(* IEC 61131-3 sources: daoli-st-library/DL_Motion (part 16) *)

(* ---- FB_DL_ResolverAngleTrackObs.st ---- *)
(* ===========================================================================
   组件名   : FB_DL_ResolverAngleTrackObs
   分类     : DL_Motion / 旋转变压器角度跟踪观测器
   一句话   : 二阶跟踪环由 sin/cos 直接跟踪角度与转速，无需反三角运算且天然解卷绕
   复杂度   : 3        版本 : v1.0.0        日期 : 2026-11-24
   开源溯源 : 无（clean-room 自研，未借鉴任何开源实现）
   输入契约 : fSin/fCos 两路瞬时值 [V]；fKp 角度环增益 [1/s]；fKi 速度环增益 [1/s²]
              fDtSec 采样周期 [s]；fAmpMin 最小有效幅值 [V]；fSpeedMax 转速限幅 [rad/s]
              fLockBand 锁定判定带宽（归一化误差） | lock band
   输出契约 : fAngleEst 跟踪角 [rad] 0..2π；fSpeedEst 跟踪转速 [rad/s]
              fErrorNorm 归一化角度误差（≈sin(θin−θest)） | normalized angle error
              xLocked 已锁定；xValid 输入有效；eStateOut 状态观测
   修改记录 : v1.0.0 2026-11-24 初版
   =========================================================================== *)

TYPE E_DL_TrackState :
(
    eTrackInit := 0,     // 初始化（粗定位） | init by coarse seed
    eTracking := 1,      // 正常跟踪 | normal tracking
    eSignalLost := 2     // 信号丢失冻结 | signal lost freeze
);
END_TYPE

FUNCTION_BLOCK FB_DL_ResolverAngleTrackObs
VAR_INPUT
    fSin : REAL;                        // 正弦路瞬时值 [V] | sine channel value [V]
    fCos : REAL;                        // 余弦路瞬时值 [V] | cosine channel value [V]
    fKp : REAL := 60.0;                 // 角度环增益 [1/s] | angle loop gain [1/s]
    fKi : REAL := 2000.0;               // 速度环增益 [1/s²] | speed loop gain [1/s^2]
    fDtSec : REAL := 0.0001;            // 采样周期 [s] | sample period [s]
    fAmpMin : REAL := 0.5;              // 最小有效幅值 [V] | minimum valid amplitude [V]
    fSpeedMax : REAL := 500.0;          // 转速限幅 [rad/s] | speed clamp [rad/s]
    fLockBand : REAL := 0.02;           // 锁定判定带宽（归一化） | lock band normalized
END_VAR
VAR_OUTPUT
    fAngleEst : REAL;                   // 跟踪角度 [rad] 0..2π | estimated angle [rad]
    fSpeedEst : REAL;                   // 跟踪转速 [rad/s] | estimated speed [rad/s]
    fErrorNorm : REAL;                  // 归一化角度误差 | normalized angle error
    xLocked : BOOL;                     // 已锁定标志 | locked flag
    xValid : BOOL;                      // 输入有效标志 | inputs valid flag
    eStateOut : E_DL_TrackState;        // 当前状态观测 | current state observation
END_VAR
VAR
    _eState : E_DL_TrackState := eTrackInit;  // 内部状态机状态 | internal state
    _fAngle : REAL;                     // 内部跟踪角 [rad] | internal tracked angle [rad]
    _fSpeed : REAL;                     // 内部跟踪转速 [rad/s] | internal tracked speed [rad/s]
    _fAmp : REAL;                       // 合成幅值 [V] | resultant amplitude [V]
    _fErr : REAL;                       // 原始角度误差 [V] | raw angle error [V]
    _fDt : REAL;                        // 钳位后采样周期 [s] | clamped dt [s]
    _xBad : BOOL;                       // 输入非有限标志 | not-finite flag
    _xBadPar : BOOL;                    // 参数非法标志 | invalid parameter flag
END_VAR

// ---- 非有限检测 ----
_xBad := (fSin <> fSin) OR ((fSin - fSin) <> (fSin - fSin))
      OR (fCos <> fCos) OR ((fCos - fCos) <> (fCos - fCos))
      OR (fDtSec <> fDtSec) OR ((fDtSec - fDtSec) <> (fDtSec - fDtSec));

// ---- 参数合法性 ----
_xBadPar := (fDtSec <= 0.0) OR (fAmpMin <= 0.0) OR (fSpeedMax <= 0.0)
         OR (fLockBand <= 0.0) OR (fKp < 0.0) OR (fKi < 0.0);

// ---- 周期钳位：跟踪环对步长极敏感，必须限幅 ----
_fDt := fDtSec;
IF _fDt < 0.000001 THEN
    _fDt := 0.000001;
ELSIF _fDt > 0.01 THEN
    _fDt := 0.01;
END_IF

// ---- 输出预置：角度与转速为积分状态，不做每拍清零 ----
fErrorNorm := 0.0;
xLocked := FALSE;
xValid := NOT (_xBad OR _xBadPar);

// ---- 合成幅值 ----
_fAmp := 0.0;
IF NOT _xBad THEN
    _fAmp := SQRT(fSin * fSin + fCos * fCos);
END_IF

CASE _eState OF
    eTrackInit:
        _fSpeed := 0.0;
        IF xValid AND (_fAmp >= fAmpMin) THEN
            // 粗定位种子：以 cos 符号区分半平面，跟踪环在后续拍内自动收敛
            IF fCos >= 0.0 THEN
                _fAngle := 0.0;
            ELSE
                _fAngle := 3.141592654;
            END_IF
            _eState := eTracking;
        END_IF
        fAngleEst := _fAngle;
        fSpeedEst := _fSpeed;

    eTracking:
        IF (NOT xValid) OR (_fAmp < fAmpMin) THEN
            _eState := eSignalLost;                // 幅值不足转冻结态
            fAngleEst := _fAngle;                  // 冻结输出保持最后可信值
            fSpeedEst := 0.0;
        ELSE
            // 误差：sin(θin)·cos(θest) − cos(θin)·sin(θest) = A·sin(θin−θest)
            _fErr := fSin * COS(_fAngle) - fCos * SIN(_fAngle);
            fErrorNorm := _fErr / _fAmp;           // 分母已由 fAmpMin 守卫

            // 二阶跟踪环：速度积分 + 角度积分
            _fSpeed := _fSpeed + fKi * fErrorNorm * _fDt;
            IF _fSpeed > fSpeedMax THEN
                _fSpeed := fSpeedMax;              // 转速限幅
            ELSIF _fSpeed < -fSpeedMax THEN
                _fSpeed := -fSpeedMax;
            END_IF

            _fAngle := _fAngle + (_fSpeed + fKp * fErrorNorm) * _fDt;
            IF _fAngle >= 6.283185307 THEN
                _fAngle := _fAngle - 6.283185307;  // 归一化到 0..2π
            ELSIF _fAngle < 0.0 THEN
                _fAngle := _fAngle + 6.283185307;
            END_IF

            fAngleEst := _fAngle;
            fSpeedEst := _fSpeed;
            xLocked := (ABS(fErrorNorm) < fLockBand);
        END_IF

    eSignalLost:
        fAngleEst := _fAngle;                      // 冻结保持，不按坏信号重新推断
        fSpeedEst := 0.0;
        IF xValid AND (_fAmp >= fAmpMin) THEN
            _eState := eTracking;                   // 信号恢复后从冻结角继续跟踪
        END_IF

ELSE
    _eState := eTrackInit;                          // 非法状态兜底回初始化
    fAngleEst := 0.0;
    fSpeedEst := 0.0;
    _fAngle := 0.0;
    _fSpeed := 0.0;
END_CASE

eStateOut := _eState;
END_FUNCTION_BLOCK

(* ---- FB_DL_ResolverFaultDetect.st ---- *)
(* ===========================================================================
   组件名   : FB_DL_ResolverFaultDetect
   分类     : DL_Motion / 旋转变压器故障检测
   一句话   : 断线（幅值过低）、短路（幅值过高）、失衡、相位异常四类分级检测与锁存
   复杂度   : 3        版本 : v1.0.0        日期 : 2026-11-24
   开源溯源 : 无（clean-room 自研，未借鉴任何开源实现）
   输入契约 : fSin/fCos 两路瞬时值 [V]；fAmpMin/fAmpMax 幅值上下限 [V]
              fImbLimitPct 失衡限值 [%]；fPhaseDiff 实测相位差 [rad]
              fPhaseExpected 期望相位差 [rad]；fPhaseTol 相位容差 [rad]
              tConfirmDelay 故障确认延时；xReset 复位上升沿
   输出契约 : eFaultClass 锁存故障类别；xFault 故障锁存；iFaultCode 分级码
              11/12=一级严重（断线/短路） 21/22=二级（失衡/相位） 99=未分类
              fAmplitude 合成幅值 [V]；fImbalancePct 即时失衡度 [%]；xValid 参数与输入有效
   修改记录 : v1.0.0 2026-11-24 初版
   =========================================================================== *)

TYPE E_DL_ResolverFault :
(
    eNoFault := 0,        // 无故障 | no fault
    eOpenWire := 1,       // 断线（幅值过低） | open wire, low amplitude
    eShortCircuit := 2,   // 短路（幅值过高） | short circuit, high amplitude
    eImbalanceFault := 3, // 两路失衡 | channel imbalance
    ePhaseFault := 4      // 相位异常 | phase anomaly
);
END_TYPE

FUNCTION_BLOCK FB_DL_ResolverFaultDetect
VAR_INPUT
    fSin : REAL;                       // 正弦路瞬时值 [V] | sine channel value [V]
    fCos : REAL;                       // 余弦路瞬时值 [V] | cosine channel value [V]
    fAmpMin : REAL := 0.5;             // 幅值下限（断线判据） [V] | amplitude low limit [V]
    fAmpMax : REAL := 9.0;             // 幅值上限（短路判据） [V] | amplitude high limit [V]
    fImbLimitPct : REAL := 5.0;        // 失衡限值 [%] | imbalance limit [%]
    fPhaseDiff : REAL := 0.0;          // 实测相位差 [rad] | measured phase difference [rad]
    fPhaseExpected : REAL := 0.0;      // 期望相位差 [rad] | expected phase difference [rad]
    fPhaseTol : REAL := 0.2;           // 相位容差 [rad] | phase tolerance [rad]
    tConfirmDelay : TIME := T#100MS;   // 故障确认延时 | fault confirm delay
    xReset : BOOL;                     // 故障复位上升沿 | fault reset rising edge
END_VAR
VAR_OUTPUT
    eFaultClass : E_DL_ResolverFault;  // 锁存故障类别（默认首项=无故障） | latched fault class
    xFault : BOOL;                     // 故障锁存标志 | latched fault flag
    iFaultCode : INT;                  // 分级故障码 0=无故障 | graded fault code
    fAmplitude : REAL;                 // 合成幅值 [V] | resultant amplitude [V]
    fImbalancePct : REAL;              // 即时失衡度 [%] | instantaneous imbalance [%]
    xValid : BOOL;                     // 输入与参数有效 | inputs and parameters valid
END_VAR
VAR
    _eCand : E_DL_ResolverFault := eNoFault;  // 本拍候选故障类别 | candidate fault class
    _fAbsSin : REAL;                   // 正弦绝对值 [V] | absolute sine [V]
    _fAbsCos : REAL;                   // 余弦绝对值 [V] | absolute cosine [V]
    _fMean : REAL;                     // 两路均值 [V] | mean magnitude [V]
    _fPhaseErr : REAL;                 // 相位偏差 [rad] | phase error [rad]
    _xBad : BOOL;                      // 输入非有限标志 | not-finite flag
    _xBadPar : BOOL;                   // 参数非法标志 | invalid parameter flag
    _tonConfirm : TON;                 // 确认延时定时器 | confirm delay timer
    _rtReset : R_TRIG;                 // 复位上升沿 | reset rising edge
END_VAR

// ---- 非有限检测 ----
_xBad := (fSin <> fSin) OR ((fSin - fSin) <> (fSin - fSin))
      OR (fCos <> fCos) OR ((fCos - fCos) <> (fCos - fCos))
      OR (fPhaseDiff <> fPhaseDiff) OR ((fPhaseDiff - fPhaseDiff) <> (fPhaseDiff - fPhaseDiff));

// ---- 参数合法性：上下限必须正向有序，其余限值必须为正 ----
_xBadPar := (fAmpMax <= fAmpMin) OR (fAmpMin < 0.0) OR (fImbLimitPct <= 0.0) OR (fPhaseTol <= 0.0);

// ---- 幅值与失衡度计算 ----
fAmplitude := 0.0;
fImbalancePct := 0.0;
_fAbsSin := 0.0;
_fAbsCos := 0.0;
IF NOT _xBad THEN
    fAmplitude := SQRT(fSin * fSin + fCos * fCos);
    _fAbsSin := ABS(fSin);
    _fAbsCos := ABS(fCos);
    _fMean := (_fAbsSin + _fAbsCos) * 0.5;
    IF _fMean > 0.000000001 THEN
        fImbalancePct := ABS(_fAbsSin - _fAbsCos) / _fMean * 100.0;   // 分母已守卫
    END_IF
END_IF

// ---- 相位偏差卷绕到 (−π, π] ----
_fPhaseErr := fPhaseDiff - fPhaseExpected;
IF _fPhaseErr > 1000000.0 THEN
    _fPhaseErr := 1000000.0;
ELSIF _fPhaseErr < -1000000.0 THEN
    _fPhaseErr := -1000000.0;
END_IF
_fPhaseErr := _fPhaseErr - 6.283185307 * TRUNC(_fPhaseErr / 6.283185307);
IF _fPhaseErr > 3.141592654 THEN
    _fPhaseErr := _fPhaseErr - 6.283185307;
ELSIF _fPhaseErr <= -3.141592654 THEN
    _fPhaseErr := _fPhaseErr + 6.283185307;
END_IF

xValid := NOT (_xBad OR _xBadPar);

// ---- 候选分类：四类判据互斥，且各有独立赋值语句（禁止共用枚举成员） ----
_eCand := eNoFault;
IF xValid THEN
    IF fAmplitude < fAmpMin THEN
        _eCand := eOpenWire;                       // 断线：幅值低于下限
    ELSIF fAmplitude > fAmpMax THEN
        _eCand := eShortCircuit;                   // 短路：幅值高于上限
    ELSIF fImbalancePct > fImbLimitPct THEN
        _eCand := eImbalanceFault;                 // 失衡：两路幅值差超限
    ELSIF ABS(_fPhaseErr) > fPhaseTol THEN
        _eCand := ePhaseFault;                     // 相位：偏差超出容差
    END_IF
END_IF

// ---- 确认延时定时器：无条件每周期调用 ----
_tonConfirm(IN := (_eCand <> eNoFault), PT := tConfirmDelay);
_rtReset(CLK := xReset);

// ---- 故障相回放锁存类别，不按当下输入重新推断 ----
IF xFault THEN
    _eCand := eFaultClass;
END_IF

// ---- 分级映射：一级（断线/短路）与二级（失衡/相位）各有独立码值 ----
iFaultCode := 0;
CASE _eCand OF
    eNoFault:
        iFaultCode := 0;                           // 无故障
    eOpenWire:
        iFaultCode := 11;                          // 一级：断线
    eShortCircuit:
        iFaultCode := 12;                          // 一级：短路
    eImbalanceFault:
        iFaultCode := 21;                          // 二级：失衡
    ePhaseFault:
        iFaultCode := 22;                          // 二级：相位异常
ELSE
    iFaultCode := 99;                              // 非法类别兜底
END_CASE

// ---- 锁存与唯一解除路径 ----
IF _tonConfirm.Q AND NOT xFault THEN
    eFaultClass := _eCand;                         // 锁存首次确认的类别
    xFault := TRUE;
END_IF
IF _rtReset.Q AND NOT xFault THEN
    eFaultClass := eNoFault;                       // 无故障时复位仅做清码
    iFaultCode := 0;
ELSIF _rtReset.Q AND xFault THEN
    xFault := FALSE;                               // 解除路径：复位上升沿
    eFaultClass := eNoFault;
    iFaultCode := 0;
END_IF
END_FUNCTION_BLOCK

(* ---- FB_DL_RotaryKnifeCutSyncCtrl.st ---- *)
(*
  Name: FB_DL_RotaryKnifeCutSyncCtrl
  Category: DL_Motion
  Version: 1.0.0
  Round: R89 / 2026-11-25
  开源溯源：clean-room 自研（族 运动同步控制，ST 开源生态实测 0 命中，无外部代码引入）
  功能：旋转刀同步定尺剪切：材料虚轴跟随 + 刀轴相位锁 + 剪切窗口判定，六相状态机含失步保护。
  边界条件：① 六浮点入参全部过非有限闸；配置越域即锁故障（101），虚轴增量强制置零、不推进；
            ② 相位比较一律做 ±180° 环绕归一化（NormalizeDeg180 方法），禁直接相减；
            ③ 相位锁判据：e = wrap180(刀相 − 180° − 材料相)。传动比 fSyncRatio = 1.0 时 e 恒 0；
               传动比偏离 1.0 时每刀漂移 (ratio − 1)×360°，|e| 超 fPhaseTolDeg 即失步，超 30° 锁故障（104）；
            ④ 剪切窗口按刀相相对 180° 的偏差定义，半宽 = fWindowDeg/2；窗口判据基于上一拍位置（滞后一拍）；
            ⑤ 遗留假设（R95 三句）：本件无周期引脚，虚轴积分用代理周期 DL_RKC_DT = 10 ms；
               该代理覆盖任务周期 1~20 ms；覆盖不到的区间（任务周期 < 1 ms 或 > 20 ms）由上层任务组态保证，
               并挂入编译验证债，交付前三平台各验证一次；
            ⑥ 使能撤销语义：位置量冻结保持末值（不归零），xSyncOk 置 FALSE（R191 已声明）；
            ⑦ 故障解除唯一路径：故障相内 xEnable 释放（R152），清锁存回 eIdle。
  状态机：eIdle / eHoming / eSyncWait / eSynced / eCutting / eReturn / eFault（CASE 含 ELSE 兜底）。
  量纲自证：v[m/min]×1000/60 = mm/s；mm/s × s ÷ mm = 转；转 × 360 = °。
*)
TYPE E_DL_RkcPhase :
(
    eIdle     := 0,     (* 待机：等使能沿 / Idle, waiting for enable edge *)
    eHoming   := 10,    (* 找零相：虚轴与刀轴归零 / Homing, both axes zeroed *)
    eSyncWait := 20,    (* 同步等待相：等相位锁进带 / Sync wait, phase lock in band *)
    eSynced   := 30,    (* 已同步相：等剪切窗口 / Synced, waiting cut window *)
    eCutting  := 40,    (* 剪切相：窗口内执行剪切 / Cutting inside window *)
    eReturn   := 50,    (* 返回相：离开窗口后回同步相 / Return after leaving window *)
    eFault    := 90     (* 故障相：锁存待释放 / Fault latched, awaiting release *)
);
END_TYPE

FUNCTION_BLOCK FB_DL_RotaryKnifeCutSyncCtrl
VAR_INPUT
    xEnable : BOOL;             (* 使能 [-] Enable *)
    fLineSpeedMpm : REAL;       (* 线速度 [m/min] Line speed [m/min] *)
    fCutLenMm : REAL;           (* 定尺长度（一个虚轴周期） [mm] Cut length per revolution [mm] *)
    fKnifeDiaMm : REAL;         (* 刀盘直径 [mm] Knife diameter [mm] *)
    fSyncRatio : REAL;          (* 传动比（刀轴角位移/虚轴角位移） [-] Sync ratio *)
    fWindowDeg : REAL;          (* 剪切窗口宽度 [°] Cutting window width [deg] *)
    fPhaseTolDeg : REAL;        (* 相位锁容差 [°] Phase lock tolerance [deg] *)
END_VAR
VAR_OUTPUT
    fMasterPosDeg : REAL;       (* 材料虚轴位置 [°] Master virtual axis position [deg] *)
    fSlavePosDeg : REAL;        (* 刀轴位置 [°] Knife axis position [deg] *)
    xInWindow : BOOL;           (* 处于剪切窗口 [-] Inside cutting window *)
    nCutCount : UDINT;          (* 累计剪切刀数（饱和） [刀] Cut counter, saturating *)
    xSyncOk : BOOL;             (* 相位锁成立 [-] Phase lock established *)
    xFault : BOOL;              (* 故障锁存标志 [-] Fault latched *)
    nErrCode : INT;             (* 故障码 0/101 组态/103 未同步进窗口/104 失步/105 非法相 [-] Error code *)
END_VAR
VAR
    _eState : E_DL_RkcPhase := E_DL_RkcPhase.eIdle;  (* 内部相（CASE 唯一写入目标） [-] Internal phase *)
    _bInit : BOOL := FALSE;         (* 首扫初始化标志 [-] First-scan init flag *)
    _bFaultLatch : BOOL := FALSE;   (* 故障锁存位 [-] Fault latch *)
    _bReqFault : BOOL := FALSE;     (* 单拍故障请求（段 2 预清） [-] Fault request *)
    _bCfgBad : BOOL := FALSE;       (* 配置非法当拍量 [-] Configuration bad *)
    _bInWindow : BOOL := FALSE;     (* 窗口判据当拍量 [-] In-window criterion *)
    _bSyncOk : BOOL := FALSE;       (* 相位锁当拍量 [-] Phase lock criterion *)
    _nErr : INT := 0;               (* 故障码锁存 [-] Latched error code *)
    _nReqErr : INT := 0;            (* 当拍请求码 [-] Requested error code *)
    _nCut : UDINT := 0;             (* 刀数累计锁存（饱和） [刀] Cut count latch *)
    _fMasterDeg : REAL := 0.0;      (* 虚轴位置保持量 [°] Master position hold [deg] *)
    _fSlaveDeg : REAL := 0.0;       (* 刀轴位置保持量 [°] Knife position hold [deg] *)
    _fAdvDeg : REAL := 0.0;         (* 单拍虚轴增量 [°] Master increment per scan [deg] *)
    _fBladeErr : REAL := 0.0;       (* 刀相相对窗口中心偏差（归一化） [°] Blade-to-center error [deg] *)
    _fLockErr : REAL := 0.0;        (* 相位锁误差（归一化） [°] Phase lock error [deg] *)
    rtEnable : R_TRIG;              (* 使能沿（段 1 无条件调用） / Enable edge *)
    rtWindow : R_TRIG;              (* 窗口进入沿（段 1 无条件调用） / Window entry edge *)
    tonHome : TON;                  (* 找零窗（段 1 无条件调用） / Homing window *)
END_VAR
VAR CONSTANT
    DL_RKC_DT : REAL := 0.01;           (* 代理扫描周期（遗留假设见头注释） [s] Proxy scan cycle [s] *)
    DL_RKC_MMPM : REAL := 1000.0;       (* 米 → 毫米换算 [mm/m] Metre to millimetre *)
    DL_RKC_SECMIN : REAL := 60.0;       (* 每秒 → 每分钟换算 [s/min] Second to minute *)
    DL_RKC_FULL : REAL := 360.0;        (* 整转角度 [°] Full revolution [deg] *)
    DL_RKC_HALF : REAL := 180.0;        (* 半转角度 [°] Half revolution [deg] *)
    DL_RKC_CUT_CENTER : REAL := 180.0;  (* 窗口中心刀相 [°] Window center blade phase [deg] *)
    DL_RKC_EXIT_MARGIN : REAL := 5.0;   (* 出窗裕度（防抖） [°] Window exit margin [deg] *)
    DL_RKC_ERR_MAX : REAL := 30.0;      (* 失步门限 [°] Loss-of-sync threshold [deg] *)
    DL_RKC_HOME : TIME := T#500MS;      (* 找零窗（确定性时窗） [ms] Homing window [ms] *)
    DL_RKC_CUT_MAX : UDINT := 4294967295;   (* 刀数饱和上限 [刀] Cut count ceiling *)
    DL_V_MIN : REAL := 0.0;             (* 线速度下限 [m/min] Line speed floor [m/min] *)
    DL_V_MAX : REAL := 600.0;           (* 线速度上限 [m/min] Line speed ceiling [m/min] *)
    DL_L_MIN : REAL := 50.0;            (* 定尺下限 [mm] Cut length floor [mm] *)
    DL_L_MAX : REAL := 20000.0;         (* 定尺上限 [mm] Cut length ceiling [mm] *)
    DL_D_MIN : REAL := 50.0;            (* 刀径下限 [mm] Knife diameter floor [mm] *)
    DL_D_MAX : REAL := 2000.0;          (* 刀径上限 [mm] Knife diameter ceiling [mm] *)
    DL_R_MIN : REAL := 0.2;             (* 传动比下限 [-] Sync ratio floor *)
    DL_R_MAX : REAL := 5.0;             (* 传动比上限 [-] Sync ratio ceiling *)
    DL_W_MIN : REAL := 1.0;             (* 窗口宽度下限 [°] Window floor [deg] *)
    DL_W_MAX : REAL := 180.0;           (* 窗口宽度上限 [°] Window ceiling [deg] *)
    DL_TOL_MIN : REAL := 0.1;           (* 相位容差下限 [°] Tolerance floor [deg] *)
    DL_TOL_MAX : REAL := 20.0;          (* 相位容差上限 [°] Tolerance ceiling [deg] *)
END_VAR

(*-----------------------------------------------------------------------------
  方法 NormalizeDeg180：把任意角度归一到 (-180, 180] 区间（±180° 环绕归一化）
  契约：入参 fDegIn [°]；返回归一化角度 [°]。非有限入参返回哨兵 0（R81 还原方向不饱和）。
  实现：三段条件减法覆盖 [-540, 540) 全域；本件两轴位置均按 [0,360) 维持，差值必落该域内，
        故无需循环，无死循环风险（R4 循环守卫结构性免除）。
-----------------------------------------------------------------------------*)
METHOD PUBLIC NormalizeDeg180 : REAL
VAR_INPUT
    fDegIn : REAL;      (* 待归一化角度 [°] Angle to normalize [deg] *)
END_VAR
VAR
    fVal : REAL := 0.0; (* 归一化中间量 [°] Normalized scratch [deg] *)
END_VAR
NormalizeDeg180 := 0.0;                             (* 出口预置哨兵 / Preset sentinel *)
IF (fDegIn <> fDegIn) OR ((fDegIn - fDegIn) <> 0.0) THEN
    NormalizeDeg180 := 0.0;                         (* 非有限：返回哨兵 0 / Non-finite to sentinel *)
    RETURN;
END_IF
fVal := fDegIn;
IF fVal >= DL_RKC_HALF THEN
    fVal := fVal - DL_RKC_FULL;                     (* 上半周折回 / Fold upper half *)
END_IF
IF fVal < (0.0 - DL_RKC_HALF) THEN
    fVal := fVal + DL_RKC_FULL;                     (* 下半周折回 / Fold lower half *)
END_IF
IF fVal >= DL_RKC_HALF THEN
    fVal := fVal - DL_RKC_FULL;                     (* 二次折回（差域上限） / Second fold *)
END_IF
NormalizeDeg180 := fVal;
END_METHOD

(* —— 段 0：非有限闸 + 虚轴增量派生 + 相位量与窗口判据 —— *)
_bCfgBad := (fLineSpeedMpm <> fLineSpeedMpm) OR ((fLineSpeedMpm - fLineSpeedMpm) <> 0.0)
         OR (fCutLenMm <> fCutLenMm) OR ((fCutLenMm - fCutLenMm) <> 0.0)
         OR (fKnifeDiaMm <> fKnifeDiaMm) OR ((fKnifeDiaMm - fKnifeDiaMm) <> 0.0)
         OR (fSyncRatio <> fSyncRatio) OR ((fSyncRatio - fSyncRatio) <> 0.0)
         OR (fWindowDeg <> fWindowDeg) OR ((fWindowDeg - fWindowDeg) <> 0.0)
         OR (fPhaseTolDeg <> fPhaseTolDeg) OR ((fPhaseTolDeg - fPhaseTolDeg) <> 0.0)
         OR (fLineSpeedMpm < DL_V_MIN) OR (fLineSpeedMpm > DL_V_MAX)
         OR (fCutLenMm < DL_L_MIN) OR (fCutLenMm > DL_L_MAX)
         OR (fKnifeDiaMm < DL_D_MIN) OR (fKnifeDiaMm > DL_D_MAX)
         OR (fSyncRatio < DL_R_MIN) OR (fSyncRatio > DL_R_MAX)
         OR (fWindowDeg < DL_W_MIN) OR (fWindowDeg > DL_W_MAX)
         OR (fPhaseTolDeg < DL_TOL_MIN) OR (fPhaseTolDeg > DL_TOL_MAX);
(* 虚轴增量：先闸后除（fCutLenMm 为除子，配置非法时强制 0，绝不进入除法） *)
IF _bCfgBad THEN
    _fAdvDeg := 0.0;
ELSE
    _fAdvDeg := ((fLineSpeedMpm * DL_RKC_MMPM) / DL_RKC_SECMIN) * DL_RKC_DT / fCutLenMm * DL_RKC_FULL;
END_IF
(* 刀相相对窗口中心偏差：±180° 归一化（禁直接相减） *)
_fBladeErr := NormalizeDeg180(_fSlaveDeg - DL_RKC_CUT_CENTER);
(* 相位锁误差：e = wrap180(刀相 − 180° − 材料相) *)
_fLockErr := NormalizeDeg180(_fSlaveDeg - DL_RKC_CUT_CENTER - _fMasterDeg);
(* 窗口判据：偏差绝对值不超过半窗宽 *)
_bInWindow := ABS(_fBladeErr) <= (fWindowDeg / 2.0);
(* 相位锁判据：误差绝对值不超容差，且已进入同步类相位 *)
_bSyncOk := (NOT _bCfgBad) AND (ABS(_fLockErr) <= fPhaseTolDeg)
            AND ((_eState = E_DL_RkcPhase.eSynced) OR (_eState = E_DL_RkcPhase.eCutting)
              OR (_eState = E_DL_RkcPhase.eReturn));
(* —— 段 1：两沿与找零 TON 无条件周期刷新（R7），禁放入分支 —— *)
rtEnable(CLK := xEnable);                                           (* 使能沿 / Enable edge *)
rtWindow(CLK := _bInWindow);                                        (* 窗口进入沿 / Window edge *)
tonHome(IN := (_eState = E_DL_RkcPhase.eHoming), PT := DL_RKC_HOME);(* 找零窗 / Homing window *)
(* —— 段 2：单拍量预清零（不含锁存/累计量，R107） —— *)
_bReqFault := FALSE;
_nReqErr := 0;
IF _bCfgBad THEN
    _bReqFault := TRUE; _nReqErr := 101;    (* 组态非法 / Configuration bad *)
END_IF
(* 首扫初始化：位置与刀数一次性归零（R310） *)
IF NOT _bInit THEN
    _fMasterDeg := 0.0;
    _fSlaveDeg := 0.0;
    _nCut := 0;
    _bInit := TRUE;
END_IF
(* —— 段 3：失步监控（同步类相位内 |e| 超门限即请求故障） —— *)
IF ((_eState = E_DL_RkcPhase.eSynced) OR (_eState = E_DL_RkcPhase.eCutting)
    OR (_eState = E_DL_RkcPhase.eReturn)) AND (ABS(_fLockErr) > DL_RKC_ERR_MAX) THEN
    _bReqFault := TRUE; _nReqErr := 104;    (* 失步 / Loss of sync *)
END_IF
(* —— 段 4：故障锁存解除（唯一路径 = 故障相内 xEnable 释放，R152） —— *)
IF _bFaultLatch AND (NOT xEnable) THEN
    _bFaultLatch := FALSE;                  (* 清锁存 / Clear latch *)
    _nErr := 0;                             (* 清码 / Clear code *)
    _eState := E_DL_RkcPhase.eIdle;         (* 迁回待机 / Back to idle *)
END_IF
(* —— 段 5：主状态机（ENUM + CASE，ELSE 兜底） —— *)
CASE _eState OF
E_DL_RkcPhase.eIdle:
    IF rtEnable.Q AND (NOT _bFaultLatch) THEN
        _fMasterDeg := 0.0;                 (* 虚轴归零 / Master zeroed *)
        _fSlaveDeg := 0.0;                  (* 刀轴归零 / Knife zeroed *)
        _nCut := 0;                         (* 刀数清零 / Cut count reset *)
        _eState := E_DL_RkcPhase.eHoming;   (* → 找零相 / To homing *)
    END_IF
E_DL_RkcPhase.eHoming:
    _fMasterDeg := _fMasterDeg + _fAdvDeg;  (* 找零期虚轴空推（材料已走） / Master advances *)
    _fSlaveDeg := _fSlaveDeg + (_fAdvDeg * fSyncRatio);   (* 刀轴按传动比跟随 / Knife follows ratio *)
    IF tonHome.Q THEN
        _eState := E_DL_RkcPhase.eSyncWait; (* 找零窗到 → 同步等待 / Home done, sync wait *)
    END_IF
E_DL_RkcPhase.eSyncWait:
    _fMasterDeg := _fMasterDeg + _fAdvDeg;  (* 虚轴推进 / Master advance *)
    _fSlaveDeg := _fSlaveDeg + (_fAdvDeg * fSyncRatio);   (* 刀轴跟随 / Knife advance *)
    IF ABS(_fLockErr) <= fPhaseTolDeg THEN
        _eState := E_DL_RkcPhase.eSynced;   (* 相位进带 → 已同步 / In band, synced *)
    END_IF
E_DL_RkcPhase.eSynced:
    _fMasterDeg := _fMasterDeg + _fAdvDeg;
    _fSlaveDeg := _fSlaveDeg + (_fAdvDeg * fSyncRatio);
    IF rtWindow.Q AND _bSyncOk THEN
        IF _nCut < DL_RKC_CUT_MAX THEN
            _nCut := _nCut + 1;             (* 刀数推进（容量载体判上限） / Saturating cut count *)
        END_IF
        _eState := E_DL_RkcPhase.eCutting;  (* → 剪切相 / To cutting *)
    ELSIF rtWindow.Q THEN
        _bReqFault := TRUE;                 (* 未同步即到切点：拒切并报失步 / Cut rejected *)
        _nReqErr := 103;
    END_IF
E_DL_RkcPhase.eCutting:
    _fMasterDeg := _fMasterDeg + _fAdvDeg;
    _fSlaveDeg := _fSlaveDeg + (_fAdvDeg * fSyncRatio);
    IF NOT _bInWindow THEN
        _eState := E_DL_RkcPhase.eReturn;   (* 出窗 → 返回相 / Window left, return *)
    END_IF
E_DL_RkcPhase.eReturn:
    _fMasterDeg := _fMasterDeg + _fAdvDeg;
    _fSlaveDeg := _fSlaveDeg + (_fAdvDeg * fSyncRatio);
    IF ABS(_fBladeErr) >= ((fWindowDeg / 2.0) + DL_RKC_EXIT_MARGIN) THEN
        _eState := E_DL_RkcPhase.eSynced;   (* 越出裕度 → 回同步相 / Past margin, synced *)
    END_IF
E_DL_RkcPhase.eFault:
    _fAdvDeg := 0.0;                        (* 故障相：虚轴增量清零，轴停在末位 / Axes hold *)
ELSE
    _bReqFault := TRUE;                     (* 非法相兜底 / Illegal phase fallback *)
    _nReqErr := 105;
END_CASE
(* 使能撤销：非故障相回待机，位置冻结保持（R191 已声明） *)
IF (NOT xEnable) AND (_eState <> E_DL_RkcPhase.eFault) AND (_eState <> E_DL_RkcPhase.eIdle) THEN
    _eState := E_DL_RkcPhase.eIdle;
END_IF
(* 位置环绕归一：两轴保持 [0,360)，防长时运行精度流失 *)
IF _fMasterDeg >= DL_RKC_FULL THEN
    _fMasterDeg := _fMasterDeg - DL_RKC_FULL;
END_IF
IF _fMasterDeg < 0.0 THEN
    _fMasterDeg := _fMasterDeg + DL_RKC_FULL;
END_IF
IF _fSlaveDeg >= DL_RKC_FULL THEN
    _fSlaveDeg := _fSlaveDeg - DL_RKC_FULL;
END_IF
IF _fSlaveDeg < 0.0 THEN
    _fSlaveDeg := _fSlaveDeg + DL_RKC_FULL;
END_IF
(* —— 段 6：故障请求统一落地（唯一锁存点 + 同步迁相，R187/R252） —— *)
IF _bReqFault AND (NOT _bFaultLatch) THEN
    _bFaultLatch := TRUE;                   (* 锁存 / Latch *)
    _nErr := _nReqErr;                      (* 码锁存回放 / Latched code *)
    _eState := E_DL_RkcPhase.eFault;        (* 同步迁相 / Migrate to fault *)
END_IF
(* —— 段 7：统一出口（各出口单点赋值） —— *)
fMasterPosDeg := _fMasterDeg;
fSlavePosDeg := _fSlaveDeg;
xInWindow := _bInWindow AND (NOT _bFaultLatch);
nCutCount := _nCut;
xSyncOk := _bSyncOk AND (NOT _bFaultLatch);
xFault := _bFaultLatch;
nErrCode := _nErr;
END_FUNCTION_BLOCK

(* ---- FB_DL_RtcpFiveAxisSeq.st ---- *)
(* ============================================================
   DL_Motion / FB_DL_RtcpFiveAxisSeq ｜ v1.0.0 ｜ 2026-11-25
   功能：五轴 RTCP 补偿相序机：eIdle → ePivotCal（摆角稳定窗 200ms + 超时狗 5s）
         → eEnable（摆角软限位校验）→ eInterp（插补补偿）→ eExit（补偿斜坡回 0）→ eIdle；
         软限位越界/补偿越限/非有限/标定超时/非法相位一律 eFault 锁存并回放码。
   边界：① 故障唯一解除 = bReset 上升沿（R152 可达）；② bReset 作用域三项：
         清锁存、迁 eIdle、清累计量与快照（不动 _bInit）；③ bEnable=FALSE 语义 =
         降级为安全值 + 置标志（经 eExit 退补到 0，非冻结保持，R191/N2）；
         ④ 同拍双窗配比：tCalTmo(5s) > tCalSettle(200ms)（R100）；
         ⑤ 出口补偿量非有限即写 0，禁 NaN 直穿 REAL（N1）。
   依赖：仅 IEC 61131-3（TON/R_TRIG/SIN/COS/ABS/MIN/MAX/LIMIT）
   溯源：DLF-A-RTCP（内部原创线）｜枚举归属：E_DL_RtcpSeqPhase 唯一属主（R264）
   码位：零 16# 范式；uErrId 0 无 / 1 组态 / 2 非有限 / 3 软限位 / 4 补偿越限 /
         5 标定超时 / 6 非法相位（码 1 含 nAxisMode ≠ 0 即工件坐标模式未实现）
   ============================================================ *)
TYPE E_DL_RtcpSeqPhase :
(
    eIdle     := 0,    // 待机：补偿关闭 / Idle with compensation off
    ePivotCal := 10,   // 枢轴标定：稳定窗 + 超时狗 / Pivot calibration window
    eEnable   := 20,   // 使能确认：软限位校验 / Enable confirmation with soft limits
    eInterp   := 30,   // 插补补偿：逐拍输出并监视越限 / Compensation output with overrun watch
    eExit     := 40,   // 退出：补偿斜坡回 0 / Exit ramp back to zero
    eFault    := 90    // 故障：锁存至复位沿 / Fault latched until the reset edge
);
END_TYPE

FUNCTION_BLOCK FB_DL_RtcpFiveAxisSeq
VAR_INPUT
    bEnable     : BOOL;   // 补偿使能电平，FALSE 触发退补 [-] / Compensation enable level
    bReset      : BOOL;   // 故障复位，上升沿解除锁存 [-] / Fault reset on the rising edge
    fPivotLenMm : REAL;   // 枢轴长度 [mm] / Pivot length in millimeters
    fTiltADeg   : REAL;   // 摆动轴 A 角反馈 [deg] / Swivel axis A angle feedback
    fTiltBDeg   : REAL;   // 摆动轴 B 角反馈 [deg] / Swivel axis B angle feedback
    nAxisMode   : DINT;   // 五轴模式 0=刀尖跟随（本件已实现）/ 1=工件坐标（未实现，判组态非法）[-] / Five axis mode selector
END_VAR
VAR_OUTPUT
    bCompActive : BOOL;   // 补偿生效（仅插补相）[-] / Compensation active in the interpolation phase
    bError      : BOOL;   // 故障锁存标志 [-] / Latched fault flag
    fCompZmm    : REAL;   // Z 向补偿量本拍生效值 [mm] / Z compensation amount in effect
    uErrId      : UDINT;  // 事件码锁存值，0 = 无事件 [-] / Latched event code
    nPhase      : INT;    // 相位号镜像 0/10/20/30/40/90 [-] / Phase number mirror
END_VAR
VAR
    rtReset      : R_TRIG;                                        // 复位沿实例，段 0 无条件刷新 / Reset edge
    tonCalSettle : TON;                                           // 标定稳定窗，段 0 无条件刷新 / Settle window
    tonCalTmo    : TON;                                           // 标定超时狗，段 0 无条件刷新 / Timeout watchdog
    _eState      : E_DL_RtcpSeqPhase := E_DL_RtcpSeqPhase.eIdle;  // 内部相位 / Internal phase
    _bInit       : BOOL := FALSE;                                 // 首扫初始化已执行 [-] / First scan init done
    _bFault      : BOOL := FALSE;                                 // 故障锁存位 [-] / Latched fault bit
    _uFault      : UDINT := 0;                                    // 故障码锁存 [-] / Latched fault code
    _bCfgBad     : BOOL;                                          // 组态非法当拍量 [-] / Illegal configuration flag
    _bNonFin     : BOOL;                                          // 入参非有限当拍量 [-] / Non-finite argument flag
    _bAngSeen    : BOOL := FALSE;                                 // 摆角前值已建立 [-] / Angle snapshot established
    _bAngStable  : BOOL := FALSE;                                 // 本拍摆角稳定 [-] / Angles stable this scan
    _fAPrev      : REAL := 0.0;                                   // 上拍 A 角快照 [deg] / Previous A snapshot
    _fBPrev      : REAL := 0.0;                                   // 上拍 B 角快照 [deg] / Previous B snapshot
    _fCompZ      : LREAL := 0.0;                                  // Z 向补偿量内部值 [mm] / Internal Z compensation
END_VAR
VAR CONSTANT
    DL_RTCP_SOFTLIM : LREAL := 110.0;                // 摆角软限位 [deg] / Soft limit of the swivel angle
    DL_RTCP_COMPLIM : LREAL := 50.0;                 // 补偿量硬限 [mm] / Hard limit of the compensation
    DL_RTCP_RAMP    : LREAL := 5.0;                  // 退补斜坡每拍步长 [mm/拍] / Exit ramp step
    DL_RTCP_STABLEPS : REAL := 0.05;                 // 摆角稳定判据带 [deg] / Angle stability tolerance
    DL_RTCP_T_SETTLE : TIME := T#200MS;              // 稳定窗时长 [ms] / Settle window duration
    DL_RTCP_T_CAL    : TIME := T#5S;                 // 标定相超时 [ms] / Calibration timeout
    DL_RTCP_C_CFG    : UDINT := 1;                   // 码 1：组态非法 / Code one, illegal configuration
    DL_RTCP_C_FIN    : UDINT := 2;                   // 码 2：入参非有限 / Code two, non-finite argument
    DL_RTCP_C_SOFT   : UDINT := 3;                   // 码 3：超软限位 / Code three, soft limit violated
    DL_RTCP_C_COMP   : UDINT := 4;                   // 码 4：补偿越限 / Code four, compensation overrun
    DL_RTCP_C_TMO    : UDINT := 5;                   // 码 5：标定超时 / Code five, calibration timeout
    DL_RTCP_C_ILL    : UDINT := 6;                   // 码 6：非法相位 / Code six, illegal phase fallback
END_VAR

(* 方法 CalcPivotComp：求 Z 向补偿量并做软限位判定；返回 TRUE = 可信。
   方法内不驻留跨拍状态，入参全经引脚传入（R3 方法设计准则）。 *)
METHOD CalcPivotComp : BOOL
VAR_INPUT
    fLenMm : REAL;   // 枢轴长度 [mm] / Pivot length
    fADeg  : REAL;   // 摆动轴 A 角 [deg] / Swivel axis A angle
    fBDeg  : REAL;   // 摆动轴 B 角 [deg] / Swivel axis B angle
END_VAR
VAR_IN_OUT
    fZmm   : LREAL;  // 计算所得 Z 补偿量（本方法写回）[mm] / Computed Z compensation written back
END_VAR
VAR
    _fAr : LREAL;  // A 角弧度 [rad] / Angle A in radians
    _fBr : LREAL;  // B 角弧度 [rad] / Angle B in radians
    _fCz : LREAL;  // Z 投影 = L×(cosA·cosB − 1) [mm] / Z projection of the pivot offset
END_VAR
VAR CONSTANT
    DL_M_PI     : LREAL := 3.14159265358979324;  // 圆周率（全精度）[-] / Pi at full precision
    DL_M_SOFT   : LREAL := 110.0;                // 摆角软限位 [deg] / Soft limit of the swivel angle
END_VAR

CalcPivotComp := FALSE;  fZmm := 0.0;            // 出口先落安全值
IF (fADeg <> fADeg) OR (fBDeg <> fBDeg) OR (fLenMm <> fLenMm)
   OR ((fLenMm - fLenMm) <> (fLenMm - fLenMm)) THEN
    RETURN;
END_IF
IF fLenMm <= 0.0 THEN RETURN; END_IF             // 组态域闸
IF (ABS(fADeg) > LREAL_TO_REAL(DL_M_SOFT)) OR (ABS(fBDeg) > LREAL_TO_REAL(DL_M_SOFT)) THEN
    RETURN;                                      // 软限位用原始角度判定（禁先夹后判）
END_IF
_fAr := REAL_TO_LREAL(fADeg) * DL_M_PI / 180.0;
_fBr := REAL_TO_LREAL(fBDeg) * DL_M_PI / 180.0;
_fCz := REAL_TO_LREAL(fLenMm) * (COS(_fAr) * COS(_fBr) - 1.0);
IF (_fCz <> _fCz) OR ((_fCz - _fCz) <> (_fCz - _fCz)) THEN
    fZmm := 0.0;  RETURN;
END_IF
fZmm := _fCz;                                     // 原值回传，越限判定归主体（保码 4 可达）
CalcPivotComp := TRUE;
END_METHOD

(* 段 0：沿实例与定时器无条件每拍刷新（R7） *)
rtReset (CLK := bReset);
tonCalSettle (IN := (_eState = E_DL_RtcpSeqPhase.ePivotCal) AND _bAngStable AND (NOT _bFault),
              PT := DL_RTCP_T_SETTLE);
tonCalTmo (IN := (_eState = E_DL_RtcpSeqPhase.ePivotCal) AND (NOT _bFault), PT := DL_RTCP_T_CAL);

(* 段 1：单拍量预清零（锁存量与快照不入清单，R107） *)
_bCfgBad := FALSE;  _bNonFin := FALSE;  _bAngStable := FALSE;

(* 段 2：首扫与复位沿同款初始化（作用域：清锁存/迁相位/清累计与快照，R310/R311） *)
IF (NOT _bInit) OR rtReset.Q THEN
    _bInit := TRUE;  _bFault := FALSE;  _uFault := 0;
    _fCompZ := 0.0;  _fAPrev := 0.0;  _fBPrev := 0.0;  _bAngSeen := FALSE;
    _eState := E_DL_RtcpSeqPhase.eIdle;
END_IF

(* 段 3：组态闸与非有限闸（覆盖全部参与换算的引脚，R272）
   模式引脚参与判据：本件换算 = A+B 双摆动 Z 投影（模式 0 刀尖跟随）；模式 1 工件坐标
   的换算分支本轮未实现，判组态非法并置码 1——禁「入闸不换算」的死引脚与两模式同形输出
   （R190 归因唯一，禁静默给出位形相同的补偿量） *)
IF (fPivotLenMm <= 0.0) OR (nAxisMode <> 0) THEN
    _bCfgBad := TRUE;
END_IF
IF (fPivotLenMm <> fPivotLenMm) OR (fTiltADeg <> fTiltADeg) OR (fTiltBDeg <> fTiltBDeg)
   OR ((fPivotLenMm - fPivotLenMm) <> (fPivotLenMm - fPivotLenMm))
   OR ((fTiltADeg - fTiltADeg) <> (fTiltADeg - fTiltADeg))
   OR ((fTiltBDeg - fTiltBDeg) <> (fTiltBDeg - fTiltBDeg)) THEN
    _bNonFin := TRUE;
END_IF

(* 段 4：摆角稳定判据与快照（快照与锁存同寿命，复位沿清零） *)
IF _bAngSeen AND (NOT _bNonFin)
   AND (ABS(fTiltADeg - _fAPrev) <= DL_RTCP_STABLEPS)
   AND (ABS(fTiltBDeg - _fBPrev) <= DL_RTCP_STABLEPS) THEN
    _bAngStable := TRUE;
END_IF
IF NOT _bNonFin THEN
    _fAPrev := fTiltADeg;  _fBPrev := fTiltBDeg;  _bAngSeen := TRUE;   // 唯一写入点
END_IF

(* 段 5：主状态机（六相全覆盖 + ELSE 非法相位兜底） *)
CASE _eState OF

E_DL_RtcpSeqPhase.eIdle:
    _fCompZ := 0.0;
    (* 非有限与组态非法分别归因（R190：成因与码一一对应，禁共码） *)
    IF _bNonFin THEN
        _bFault := TRUE;  _uFault := DL_RTCP_C_FIN;  _eState := E_DL_RtcpSeqPhase.eFault;
    ELSIF _bCfgBad THEN
        _bFault := TRUE;  _uFault := DL_RTCP_C_CFG;  _eState := E_DL_RtcpSeqPhase.eFault;
    ELSIF bEnable AND (NOT _bFault) THEN
        _eState := E_DL_RtcpSeqPhase.ePivotCal;      // 拍 N+1 转出到标定相
    END_IF

E_DL_RtcpSeqPhase.ePivotCal:
    IF _bNonFin THEN
        _bFault := TRUE;  _uFault := DL_RTCP_C_FIN;  _eState := E_DL_RtcpSeqPhase.eFault;
    ELSIF _bCfgBad THEN
        _bFault := TRUE;  _uFault := DL_RTCP_C_CFG;  _eState := E_DL_RtcpSeqPhase.eFault;
    ELSIF NOT bEnable THEN
        _eState := E_DL_RtcpSeqPhase.eExit;          // 撤能使：不驻留标定相
    ELSIF tonCalTmo.Q THEN
        _bFault := TRUE;  _uFault := DL_RTCP_C_TMO;  _eState := E_DL_RtcpSeqPhase.eFault;
    ELSIF tonCalSettle.Q THEN
        _eState := E_DL_RtcpSeqPhase.eEnable;        // 拍 N+1 转出：标定完成
    END_IF

E_DL_RtcpSeqPhase.eEnable:
    (* 迁入执行相前的全量闸位复检（R274）：非有限与组态非法分别归因，禁误归软限位码 3 *)
    IF _bNonFin THEN
        _fCompZ := 0.0;  _bFault := TRUE;  _uFault := DL_RTCP_C_FIN;
        _eState := E_DL_RtcpSeqPhase.eFault;
    ELSIF _bCfgBad THEN
        _bFault := TRUE;  _uFault := DL_RTCP_C_CFG;
        _eState := E_DL_RtcpSeqPhase.eFault;
    ELSIF ABS(fTiltADeg) > LREAL_TO_REAL(DL_RTCP_SOFTLIM) THEN
        _bFault := TRUE;  _uFault := DL_RTCP_C_SOFT;  _eState := E_DL_RtcpSeqPhase.eFault;
    ELSIF ABS(fTiltBDeg) > LREAL_TO_REAL(DL_RTCP_SOFTLIM) THEN
        _bFault := TRUE;  _uFault := DL_RTCP_C_SOFT;  _eState := E_DL_RtcpSeqPhase.eFault;
    ELSIF NOT bEnable THEN
        _eState := E_DL_RtcpSeqPhase.eExit;
    ELSE
        _eState := E_DL_RtcpSeqPhase.eInterp;        // 迁入执行相：闸位已全量复检（R274）
    END_IF

E_DL_RtcpSeqPhase.eInterp:
    IF NOT bEnable THEN
        _eState := E_DL_RtcpSeqPhase.eExit;
    ELSIF _bNonFin THEN
        _fCompZ := 0.0;  _bFault := TRUE;  _uFault := DL_RTCP_C_FIN;
        _eState := E_DL_RtcpSeqPhase.eFault;
    ELSIF _bCfgBad THEN
        _fCompZ := 0.0;  _bFault := TRUE;  _uFault := DL_RTCP_C_CFG;
        _eState := E_DL_RtcpSeqPhase.eFault;         // 运行中组态非法（模式改号）：独立归因
    ELSIF NOT CalcPivotComp(fLenMm := fPivotLenMm, fADeg := fTiltADeg, fBDeg := fTiltBDeg, fZmm := _fCompZ) THEN
        _fCompZ := 0.0;  _bFault := TRUE;  _uFault := DL_RTCP_C_SOFT;
        _eState := E_DL_RtcpSeqPhase.eFault;         // 方法拒收：归因软限位
    ELSIF ABS(_fCompZ) > DL_RTCP_COMPLIM THEN
        _fCompZ := 0.0;  _bFault := TRUE;  _uFault := DL_RTCP_C_COMP;
        _eState := E_DL_RtcpSeqPhase.eFault;         // 补偿越限：独立归因（R190）
    END_IF

E_DL_RtcpSeqPhase.eExit:
    IF _fCompZ > 0.0 THEN
        _fCompZ := MAX(0.0, _fCompZ - DL_RTCP_RAMP);
    ELSIF _fCompZ < 0.0 THEN
        _fCompZ := MIN(0.0, _fCompZ + DL_RTCP_RAMP);
    ELSE
        _fCompZ := 0.0;  _eState := E_DL_RtcpSeqPhase.eIdle;   // 补偿归零才迁出
    END_IF

E_DL_RtcpSeqPhase.eFault:
    _fCompZ := 0.0;                                              // 故障相：补偿压 0（N1/N3）
    IF rtReset.Q THEN _eState := E_DL_RtcpSeqPhase.eIdle; END_IF // 唯一解除路径

ELSE
    _bFault := TRUE;  _uFault := DL_RTCP_C_ILL;  _eState := E_DL_RtcpSeqPhase.eFault;
END_CASE

(* 段 6：故障迁相闸（置于解除段之后，R274） *)
IF _bFault AND (_eState <> E_DL_RtcpSeqPhase.eFault) THEN
    _eState := E_DL_RtcpSeqPhase.eFault;
END_IF

(* 段 7：统一出口段（判据位与实值单点裁决，N4/R191） *)
bCompActive := (_eState = E_DL_RtcpSeqPhase.eInterp);
bError := _bFault;  uErrId := _uFault;
IF (_eState = E_DL_RtcpSeqPhase.eInterp) AND (_fCompZ = _fCompZ)
   AND ((_fCompZ - _fCompZ) = (_fCompZ - _fCompZ)) THEN
    fCompZmm := LREAL_TO_REAL(_fCompZ);
ELSE
    fCompZmm := 0.0;                                            // 非插补相或非有限：落 0（N1）
END_IF

(* 相位号镜像：单一 CASE 映射，禁多分支重复写同一状态（R20） *)
CASE _eState OF
    E_DL_RtcpSeqPhase.eIdle:     nPhase := 0;
    E_DL_RtcpSeqPhase.ePivotCal: nPhase := 10;
    E_DL_RtcpSeqPhase.eEnable:   nPhase := 20;
    E_DL_RtcpSeqPhase.eInterp:   nPhase := 30;
    E_DL_RtcpSeqPhase.eExit:     nPhase := 40;
    E_DL_RtcpSeqPhase.eFault:    nPhase := 90;
ELSE
    nPhase := 90;
END_CASE
END_FUNCTION_BLOCK

(* ---- FB_DL_ScreenPrintAlign.st ---- *)
// =====================================================================
// FB_DL_ScreenPrintAlign.st
// 丝网印刷对位（相机 dx/dy/dθ → XY 纠偏相对定位 → 公差判定）
// Screen printing alignment FB via I_DL_MotionAxis contract
// 码位: 16#0004_0340 ~ 16#0004_0344 (本件独占 5 槽)
// 修改记录: R29 初版 (按 DISPATCH_R29 序 12)
// =====================================================================
// 枚举: E_DL_ScreenPrintState（归属 Ownership：E_DL_ScreenPrintState 归属本文件
//       FB_DL_ScreenPrintAlign，全库唯一定义，本件只定义不重声明）
//       R74 说明：本件原借用 DL_Motion/FB_DL_StringCutAlign 的 E_DL_ScreenPrintState，
//       该枚举成员集为 ( eIdle/eCalc/eWaitPos/eDone/eFault )，无 eMove 与 eVerify，
//       跨件借用即产生 E048 未解析引用；两件相位语义域不同（本件为相机对位四相），
//       故按 R264 归属断言改为携带自有枚举，成员集按本文件实际用到的相位取值。
// =====================================================================
TYPE E_DL_ScreenPrintState :
(
    eIdle   := 0,     // 空闲待触发 / Idle, waiting for trigger
    eCalc   := 10,    // 计算相：θ 补偿换算 / Calculating theta compensation
    eMove   := 20,    // 移动相：XY 逐轴相对定位 / Moving, per-axis relative positioning
    eVerify := 30,    // 验证相：公差判定 / Verifying tolerance verdict
    eDone   := 40,    // 完成态：结论保持至下一触发 / Done, verdict held until next trigger
    eFault  := 90     // 故障锁存态（仅 bReset 沿迁出）/ Fault latched, exits on reset edge
);
END_TYPE

// =====================================================================
FUNCTION_BLOCK FB_DL_ScreenPrintAlign
VAR_INPUT
    bEnable         : BOOL  := FALSE;   // 使能 / Enable
    bTrigger        : BOOL  := FALSE;   // 上升沿启动一次对位 / Trigger on rising edge
    bReset          : BOOL  := FALSE;   // 复位故障 / Reset
    fCamDx_mm       : REAL  := 0.0;     // 相机 X 偏差 -20~20 mm / Camera dX [mm]
    fCamDy_mm       : REAL  := 0.0;     // 相机 Y 偏差 -20~20 mm / Camera dY [mm]
    fCamDTheta_deg  : REAL  := 0.0;     // 相机角度偏差 -10~10 ° / Camera dTheta [deg]
    fRotRadius_mm   : REAL  := 200.0;   // 旋转补偿半径 10~2000 mm / Rotation radius [mm]
    fTol_mm         : REAL  := 0.02;    // XY 公差 0.001~2 mm / XY tolerance [mm]
    fTolTheta_deg   : REAL  := 0.05;    // 角度公差 0.001~2 ° / Theta tolerance [deg]
    fCorrMax_mm     : REAL  := 5.0;     // 最大可纠偏差 0.1~20 mm / Max correctable [mm]
    fSpeed_mmS      : REAL  := 20.0;    // 定位速度 1~200 mm/s / Speed [mm/s]
    tMoveMax        : TIME  := T#5S;    // 单次定位超时 T#100MS~T#60S / Move timeout [s]
    uRetryMax       : USINT  := 3;      // 最大重试次数 1~10 / Max retries
END_VAR
VAR_IN_OUT
    iAxisX          : I_DL_MotionAxis;  // X 轴契约引用 / X axis interface
    iAxisY          : I_DL_MotionAxis;  // Y 轴契约引用 / Y axis interface
END_VAR
VAR_OUTPUT
    fCorrX_mm       : REAL;             // 本次 X 纠偏量 mm / X correction [mm]
    fCorrY_mm       : REAL;             // 本次 Y 纠偏量 mm / Y correction [mm]
    bInTol          : BOOL;             // 纠偏后进公差 / In tolerance
    bDegraded       : BOOL;             // θ 超差不旋转降级 / Theta degraded
    uRetryCnt       : USINT;            // 已重试次数 / Retry count
    eState          : E_DL_ScreenPrintState;  // 状态 / State
    eErr            : UDINT;            // 错误码 / Error code
END_VAR
VAR
    rtrigTrigger    : R_TRIG;           // 触发沿检测（无条件刷新）/ Trigger edge detector
    fThetaRad       : REAL;             // θ 弧度值 / Theta in radians [rad]
    fCorrXTarget    : REAL;             // X 纠偏目标 / X correction target [mm]
    fCorrYTarget    : REAL;             // Y 纠偏目标 / Y correction target [mm]
    bXDone          : BOOL := FALSE;    // X 轴完成标志（换轴前清）/ X done flag, cleared on axis switch
    bXIssued        : BOOL := FALSE;    // X 轴指令已发单锁（防每拍重复下发）/ X single-shot issued lock
    bYIssued        : BOOL := FALSE;    // Y 轴指令已发单锁（防每拍重复下发）/ Y single-shot issued lock
    bAxisOk         : BOOL;             // 轴指令受理标记 / Axis command accepted
    tonMove         : TON;              // 定位超时定时器（无条件刷新）/ Move timeout timer
    tMoveMaxS       : REAL;             // 超时秒值 / Timeout seconds [s]
    xFirstScan      : BOOL  := TRUE;    // 首扫标记 / First-scan flag
END_VAR

// ---------------------------------------------------------------------
// 代码位表（本件独占，勿复用）:
//   16#0004_0340 信息 对位完成（eDone）
//   16#0004_0341 故障 偏差/参数非有限 / tMoveMax 非法 / 轴接口未就绪
//   16#0004_0342 故障 fTol_mm ≤ 0 / fSpeed_mmS ≤ 0 / uRetryMax = 0（组态错）
//   16#0004_0343 信息 ABS(fCamDTheta_deg) > fTolTheta_deg → 仅 XY 纠偏（bDegraded=TRUE）
//   16#0004_0344 故障 ABS(dx)>fCorrMax 或 ABS(dy)>fCorrMax → 拒纠；或重试达上限仍未进公差
// ---------------------------------------------------------------------

// ---- 超时秒值 / Timeout seconds ----
tMoveMaxS := TIME_TO_REAL(tMoveMax) / 1000.0;   // 秒值 / Seconds [s]

// ---- 触发沿检测（每拍无条件刷新，R7 纪律）/ Trigger edge, unconditional refresh ----
rtrigTrigger(CLK := bTrigger);  // 沿检测 / Edge detection

// ---- 非有限与时域闸 / Finite and time-domain gate ----
IF (fCamDx_mm <> fCamDx_mm) OR (ABS(fCamDx_mm) >= 1.0E12)
   OR (fCamDy_mm <> fCamDy_mm) OR (ABS(fCamDy_mm) >= 1.0E12)
   OR (fCamDTheta_deg <> fCamDTheta_deg) OR (ABS(fCamDTheta_deg) >= 1.0E12)
   OR (fRotRadius_mm <> fRotRadius_mm) OR (ABS(fRotRadius_mm) >= 1.0E12)
   OR (fTol_mm <> fTol_mm) OR (ABS(fTol_mm) >= 1.0E12)
   OR (fCorrMax_mm <> fCorrMax_mm) OR (ABS(fCorrMax_mm) >= 1.0E12)
   OR (fSpeed_mmS <> fSpeed_mmS) OR (ABS(fSpeed_mmS) >= 1.0E12)
   OR (tMoveMax = T#0MS) OR (tMoveMaxS < 0.1) OR (tMoveMaxS > 60.0) THEN
    eState := E_DL_ScreenPrintState.eFault;   // 故障态 / Fault state
    eErr := 16#0004_0341;       // 故障码 / Fault code
    RETURN;                     // 本拍结束 / End of cycle
END_IF

// ---- 组态错闸 / Configuration fault gate ----
IF (fTol_mm <= 0.0) OR (fSpeed_mmS <= 0.0) OR (uRetryMax = 0) THEN
    eState := E_DL_ScreenPrintState.eFault;   // 故障态 / Fault state
    eErr := 16#0004_0342;       // 故障码 / Fault code
    RETURN;                     // 本拍结束 / End of cycle
END_IF

// ---- 首扫初始化（R16 首扫纪律）/ First-scan initialization ----
IF xFirstScan THEN
    eState := E_DL_ScreenPrintState.eIdle;    // 空闲态 / Idle
    bInTol := FALSE;            // 结论复位 / Verdict reset
    xFirstScan := FALSE;        // 清标记 / Clear flag
END_IF

// ---- 使能撤销 / Disable ----
IF NOT bEnable THEN
    eState := E_DL_ScreenPrintState.eIdle;    // 回空闲 / Idle
    bInTol := FALSE;            // 结论复位 / Verdict reset
    bDegraded := FALSE;         // 降级复位 / Degraded reset
    uRetryCnt := 0;             // 重试清零 / Retry cleared
    RETURN;                     // 本拍结束 / End of cycle
END_IF

// ---- 故障复位 / Fault reset ----
IF (eState = E_DL_ScreenPrintState.eFault) AND bReset THEN
    eState := E_DL_ScreenPrintState.eIdle;    // 回空闲 / Idle
    uRetryCnt := 0;             // 重试清零 / Retry cleared
    bInTol := FALSE;            // 结论复位 / Verdict reset
END_IF

// ---- θ 降级判（先于状态机，供信息级登记）/ Theta degradation check ----
bDegraded := (ABS(fCamDTheta_deg) > fTolTheta_deg);     // 降级标志 / Degraded flag

// ---- 状态机 / State machine ----
CASE eState OF

    E_DL_ScreenPrintState.eIdle:      // 空闲态 / Idle
        bInTol := FALSE;        // 结论复位 / Verdict reset
        eErr := 16#0004_0340;   // 信息级：空闲正常 / Info: idle
        // 触发沿受理（bBusy 期丢弃新触发不排队）/ Accept trigger edge
        IF rtrigTrigger.Q THEN
            // 拒纠闸：偏差超最大可纠值 → 不动轴直接故障 / Reject oversize deviation
            IF (ABS(fCamDx_mm) > fCorrMax_mm) OR (ABS(fCamDy_mm) > fCorrMax_mm) THEN
                eState := E_DL_ScreenPrintState.eFault;   // 故障态 / Fault
                eErr := 16#0004_0344;   // 故障码：拒纠 / Fault: rejected
            ELSIF (iAxisX = 0) OR (iAxisY = 0) THEN    // 接口引用未注入判定（引用为空判零口径）/ Interface reference not injected, null-reference test
                eState := E_DL_ScreenPrintState.eFault;   // 故障态 / Fault
                eErr := 16#0004_0341;   // 故障码：接口未就绪 / Fault: interface
            ELSE
                eState := E_DL_ScreenPrintState.eCalc;    // 进入计算相 / Go to calc
            END_IF
        END_IF

    E_DL_ScreenPrintState.eCalc:      // 计算相：θ 补偿换算 / Calc: theta compensation
        // 小角度近似适用域注释：|θ|≤10° 内 SIN 近似线性误差 <0.5 %
        // Small-angle approximation valid for |theta| <= 10 deg, error < 0.5 %
        fThetaRad := fCamDTheta_deg * 3.14159265 / 180.0;   // 度转弧度 / Deg to rad
        // 旋转臂分解（θ 补偿项按半径投影）/ Rotational arm decomposition
        fCorrXTarget := fCamDx_mm - fThetaRad * fRotRadius_mm;  // X 目标含 θ 补偿 / X target
        fCorrYTarget := fCamDy_mm;      // Y 目标不含旋转投影 / Y target
        fCorrX_mm := fCorrXTarget;      // 输出 X 纠偏 / Output X
        fCorrY_mm := fCorrYTarget;      // 输出 Y 纠偏 / Output Y
        uRetryCnt := 0;             // 本轮重试清零 / Retry cleared
        eState := E_DL_ScreenPrintState.eMove;    // 进入移动相 / Go to move

    E_DL_ScreenPrintState.eMove:      // 移动相：单轴相对定位 / Move: relative positioning per axis
        tonMove(IN := TRUE, PT := tMoveMax);    // 超时定时器无条件刷新 / Unconditional refresh
        IF tonMove.Q THEN
            // 超时：中止不再发新指令（R27 教训）/ Timeout: abort, no new commands
            eState := E_DL_ScreenPrintState.eFault;   // 故障态 / Fault
            eErr := 16#0004_0341;   // 故障码 / Fault code
            RETURN;                 // 本拍结束 / End of cycle
        END_IF
        IF NOT bXDone THEN
            // X 轴：先发单再等到位（接口契约 MoveRelative(fDist, fVel, fAcc)，无 bDone 引脚，
            // 到位判据取 eState = eStandstill；单发语义由本件 bXIssued 单发锁承担）
            // X axis: issue once, then wait for arrival (contract has no bDone pin;
            // arrival is eState = eStandstill, single-shot owned by bXIssued)
            IF NOT bXIssued THEN
                IF iAxisX.MoveRelative(fDist := fCorrXTarget, fVel := fSpeed_mmS,
                                       fAcc := fSpeed_mmS * 10.0) THEN   // 1/10 秒达速等效加减速度 [mm/s²] / Equivalent accel
                    bXIssued := TRUE;       // 已发单 / Issued
                    bAxisOk := TRUE;        // 受理 / Accepted
                ELSE
                    eState := E_DL_ScreenPrintState.eFault;   // 指令拒绝 → 故障 / Rejected
                    eErr := 16#0004_0341;   // 故障码 / Fault code
                    RETURN;             // 本拍结束 / End of cycle
                END_IF
            ELSIF iAxisX.bError THEN
                eState := E_DL_ScreenPrintState.eFault;   // 轴错误 → 故障 / Axis error
                eErr := 16#0004_0341;   // 故障码 / Fault code
                RETURN;                 // 本拍结束 / End of cycle
            ELSIF iAxisX.eState = E_DL_AxisState.eStandstill THEN
                bXDone := TRUE;         // X 到位（待机态），换 Y 前清 X 标记（R27 教训）/ X arrived
                bXIssued := FALSE;      // 清单发锁，供 Y 轴复用 / Release single-shot
                tonMove(IN := FALSE, PT := tMoveMax);   // 重置超时 / Reset timeout
            END_IF
        ELSE
            // Y 轴：同构（契约三参数口径）/ Y axis, same three-parameter contract
            IF NOT bYIssued THEN
                IF iAxisY.MoveRelative(fDist := fCorrYTarget, fVel := fSpeed_mmS,
                                       fAcc := fSpeed_mmS * 10.0) THEN   // 等效加减速度 [mm/s²] / Equivalent accel
                    bYIssued := TRUE;       // 已发单 / Issued
                    bAxisOk := TRUE;        // 受理 / Accepted
                ELSE
                    eState := E_DL_ScreenPrintState.eFault;   // 指令拒绝 → 故障 / Rejected
                    eErr := 16#0004_0341;   // 故障码 / Fault code
                    RETURN;             // 本拍结束 / End of cycle
                END_IF
            ELSIF iAxisY.bError THEN
                eState := E_DL_ScreenPrintState.eFault;   // 轴错误 → 故障 / Axis error
                eErr := 16#0004_0341;   // 故障码 / Fault code
                RETURN;                 // 本拍结束 / End of cycle
            ELSIF iAxisY.eState = E_DL_AxisState.eStandstill THEN
                bXDone := FALSE;        // 清轴标志（换轴前清，R27 教训）/ Clear axis flag
                bYIssued := FALSE;      // 清单发锁 / Release single-shot
                eState := E_DL_ScreenPrintState.eVerify;  // 进入验证相 / Go to verify
            END_IF
        END_IF

    E_DL_ScreenPrintState.eVerify:    // 验证相：公差判定 / Verify: tolerance verdict
        // 边界含等号 / Boundary inclusive
        IF (ABS(fCamDx_mm) <= fTol_mm) AND (ABS(fCamDy_mm) <= fTol_mm) THEN
            bInTol := TRUE;     // 进公差 / In tolerance
            eState := E_DL_ScreenPrintState.eDone;    // 完成态 / Done
        ELSE
            uRetryCnt := uRetryCnt + 1;     // 重试计数 / Retry count
            IF uRetryCnt >= uRetryMax THEN
                eState := E_DL_ScreenPrintState.eFault;   // 重试耗尽 → 故障锁存 / Fault latch
                eErr := 16#0004_0344;   // 故障码 / Fault code
            ELSE
                eState := E_DL_ScreenPrintState.eMove;    // 重发定位 / Retry move
            END_IF
        END_IF

    E_DL_ScreenPrintState.eDone:      // 完成态 / Done
        bInTol := TRUE;         // 结论保持 / Verdict held
        eErr := 16#0004_0340;   // 信息级：对位完成 / Info: done
        // θ 降级信息级登记（完成且降级时覆盖信息码）/ Degraded info code
        IF bDegraded THEN
            eErr := 16#0004_0343;   // 信息级：仅 XY 纠偏 / Info: XY only
        END_IF
        // 下一触发沿重新进入计算相 / Next trigger restarts
        IF rtrigTrigger.Q THEN
            eState := E_DL_ScreenPrintState.eCalc;    // 重启 / Restart
        END_IF

    E_DL_ScreenPrintState.eFault:     // 故障态 / Fault
        bInTol := FALSE;        // 结论复位 / Verdict reset
        // eErr 已在置故障处赋值，锁存回放不重推断 / Code latched
        IF bReset THEN
            eState := E_DL_ScreenPrintState.eIdle;    // 复位回空闲 / Reset to idle
            uRetryCnt := 0;     // 重试清零 / Retry cleared
        END_IF

    ELSE                        // 非法状态拦截 / Illegal state interception
        eState := E_DL_ScreenPrintState.eFault;   // 落故障态 / Fall to fault
        eErr := 16#0004_0341;   // 故障码 / Fault code
END_CASE

// ---- 降级信息级（非完成态也登记，供上位观察）/ Degraded info outside done ----
IF bDegraded AND (eState = E_DL_ScreenPrintState.eMove) AND (eErr = 16#0004_0340) THEN
    eErr := 16#0004_0343;       // 信息级：仅 XY / Info: XY only
END_IF

END_FUNCTION_BLOCK

(* ---- FB_DL_ServoBrakeReleaseSeq.st ---- *)
(* ===========================================================================
   组件名   : FB_DL_ServoBrakeReleaseSeq
   分类     : DL_Motion / 伺服抱闸时序
   一句话   : 抱闸释放与闭合时序：先励磁后释放、先卸转矩后抱闸，含确认反馈与逐步超时
   复杂度   : 2        版本 : v1.0.0        日期 : 2026-11-24
   开源溯源 : 无（clean-room 自研，未借鉴任何开源实现）
   输入契约 : xOpenReq 释放请求；xCloseReq 闭合请求；xExciteFbk 励磁就绪反馈
              xBrakeOpenFbk 抱闸已释放反馈；xBrakeClosedFbk 抱闸已闭合反馈
              lrTorqueFbk 实际转矩反馈 [%]；lrTorqueZeroBand 零转矩判定带宽 [%]
              t*Timeout 各步超时；xReset 复位上升沿
   输出契约 : xExciteCmd 励磁指令；xBrakeReleaseCmd 抱闸释放指令 TRUE=释放
              xTorqueHoldCmd 零转矩保持指令；xOpenDone / xCloseDone 完成标志
              xError 故障锁存（唯一解除路径 = xReset 上升沿 AND 无释放请求）
              iErrorCode 1=励磁超时 2=释放超时 3=卸转矩超时 4=闭合超时 5=转矩非有限 9=非法状态
   修改记录 : v1.0.0 2026-11-24 初版
   =========================================================================== *)

TYPE E_DL_ServoBrakeState :
(
    eIdle := 0,           // 空闲 | idle
    eExcite := 1,         // 下发励磁 | issue excitation
    eWaitExcite := 2,     // 等待励磁反馈 | wait excitation feedback
    eReleaseBrake := 3,   // 下发抱闸释放 | issue brake release
    eWaitBrakeOpen := 4,  // 等待抱闸释放反馈 | wait brake open feedback
    eReady := 5,          // 释放完成保持 | release done hold
    eHoldTorque := 6,     // 卸转矩到零 | unload torque to zero
    eCloseBrake := 7,     // 下发抱闸闭合 | issue brake close
    eWaitBrakeClose := 8, // 等待抱闸闭合反馈 | wait brake close feedback
    eDone := 9,           // 闭合完成 | close done
    eFault := 10          // 故障锁存态 | latched fault
);
END_TYPE

FUNCTION_BLOCK FB_DL_ServoBrakeReleaseSeq
VAR_INPUT
    xOpenReq : BOOL;                        // 抱闸释放请求 | brake open request
    xCloseReq : BOOL;                       // 抱闸闭合请求 | brake close request
    xExciteFbk : BOOL;                      // 励磁就绪反馈 | excitation ready feedback
    xBrakeOpenFbk : BOOL;                   // 抱闸已释放反馈 | brake opened feedback
    xBrakeClosedFbk : BOOL;                 // 抱闸已闭合反馈 | brake closed feedback
    lrTorqueFbk : LREAL;                    // 实际转矩反馈 [%] | actual torque feedback [%]
    lrTorqueZeroBand : LREAL := 2.0;        // 零转矩判定带宽 [%] | zero torque band [%]
    tExciteTimeout : TIME := T#2S;          // 励磁超时 | excitation timeout
    tBrakeOpenTimeout : TIME := T#2S;       // 抱闸释放超时 | brake open timeout
    tTorqueZeroTimeout : TIME := T#5S;      // 卸转矩超时 | torque unload timeout
    tBrakeCloseTimeout : TIME := T#2S;      // 抱闸闭合超时 | brake close timeout
    xReset : BOOL;                          // 故障复位上升沿 | fault reset rising edge
END_VAR
VAR_OUTPUT
    xExciteCmd : BOOL;                      // 励磁指令 | excitation command
    xBrakeReleaseCmd : BOOL;                // 抱闸释放指令 TRUE=释放 | brake release command
    xTorqueHoldCmd : BOOL;                  // 零转矩保持指令 | zero torque hold command
    xOpenDone : BOOL;                       // 释放完成 | open done
    xCloseDone : BOOL;                      // 闭合完成 | close done
    xError : BOOL;                          // 故障锁存 | latched fault
    iErrorCode : INT;                       // 故障码 0=无故障 | error code
    eStateOut : E_DL_ServoBrakeState;         // 当前状态观测 | current state observation
END_VAR
VAR
    _eState : E_DL_ServoBrakeState := eIdle;  // 内部状态机状态 | internal state
    _xTorqueOk : BOOL;                      // 转矩已到零带内 | torque within zero band
    _tonExcite : TON;                       // 励磁等待定时器 | excitation wait timer
    _tonOpen : TON;                         // 释放等待定时器 | open wait timer
    _tonTorque : TON;                       // 卸转矩定时器 | torque unload timer
    _tonClose : TON;                        // 闭合等待定时器 | close wait timer
    _rtReset : R_TRIG;                      // 复位上升沿 | reset rising edge
END_VAR

// ---- 转矩零带判定：带宽须为正且转矩值须有限 ----
_xTorqueOk := FALSE;
IF (lrTorqueZeroBand > 0.0)
   AND NOT ((lrTorqueFbk <> lrTorqueFbk) OR ((lrTorqueFbk - lrTorqueFbk) <> (lrTorqueFbk - lrTorqueFbk)))
   AND (ABS(lrTorqueFbk) < lrTorqueZeroBand) THEN
    _xTorqueOk := TRUE;
END_IF

// ---- 定时器与边沿：无条件每周期调用 ----
_tonExcite(IN := (_eState = eWaitExcite), PT := tExciteTimeout);
_tonOpen(IN := (_eState = eWaitBrakeOpen), PT := tBrakeOpenTimeout);
_tonTorque(IN := (_eState = eHoldTorque), PT := tTorqueZeroTimeout);
_tonClose(IN := (_eState = eWaitBrakeClose), PT := tBrakeCloseTimeout);
_rtReset(CLK := xReset);

// ---- 逐拍输出预置：非锁存量复位，xError / iErrorCode 保持 ----
xExciteCmd := FALSE;
xBrakeReleaseCmd := FALSE;
xTorqueHoldCmd := FALSE;

CASE _eState OF
    eIdle:
        IF xOpenReq AND NOT xError THEN
            _eState := eExcite;
        END_IF

    eExcite:
        xExciteCmd := TRUE;                      // 先建励磁，保证抱闸打开时无溜车
        _eState := eWaitExcite;

    eWaitExcite:
        xExciteCmd := TRUE;
        IF xExciteFbk THEN
            _eState := eReleaseBrake;
        ELSIF _tonExcite.Q THEN
            xError := TRUE; iErrorCode := 1;     // 励磁超时
            _eState := eFault;
        END_IF

    eReleaseBrake:
        xExciteCmd := TRUE;
        xBrakeReleaseCmd := TRUE;                // 励磁已就绪，释放抱闸
        _eState := eWaitBrakeOpen;

    eWaitBrakeOpen:
        xExciteCmd := TRUE;
        xBrakeReleaseCmd := TRUE;
        IF xBrakeOpenFbk THEN
            _eState := eReady;
        ELSIF _tonOpen.Q THEN
            xError := TRUE; iErrorCode := 2;     // 抱闸释放超时
            _eState := eFault;
        END_IF

    eReady:
        xExciteCmd := TRUE;
        xBrakeReleaseCmd := TRUE;
        IF xCloseReq OR NOT xOpenReq THEN
            _eState := eHoldTorque;              // 收到闭合请求或撤请求，先卸转矩
        END_IF

    eHoldTorque:
        xExciteCmd := TRUE;
        xBrakeReleaseCmd := TRUE;                // 抱闸仍保持释放，仅撤转矩
        xTorqueHoldCmd := TRUE;
        IF _xTorqueOk THEN
            _eState := eCloseBrake;
        ELSIF _tonTorque.Q THEN
            xError := TRUE; iErrorCode := 3;     // 卸转矩超时
            _eState := eFault;
        END_IF

    eCloseBrake:
        xExciteCmd := TRUE;
        xTorqueHoldCmd := TRUE;
        xBrakeReleaseCmd := FALSE;               // 转矩已到零，闭合抱闸
        _eState := eWaitBrakeClose;

    eWaitBrakeClose:
        xExciteCmd := TRUE;
        xTorqueHoldCmd := TRUE;
        IF xBrakeClosedFbk THEN
            _eState := eDone;
        ELSIF _tonClose.Q THEN
            xError := TRUE; iErrorCode := 4;     // 抱闸闭合超时
            _eState := eFault;
        END_IF

    eDone:
        IF NOT xOpenReq THEN
            _eState := eIdle;                    // 请求撤销后回空闲
        END_IF

    eFault:
        xError := TRUE;                          // 故障锁存保持，抱闸因失电而夹紧
        IF _rtReset.Q AND NOT xOpenReq THEN
            xError := FALSE;                     // 唯一解除路径：复位沿且无释放请求
            iErrorCode := 0;
            _eState := eIdle;
        END_IF

ELSE
    xError := TRUE; iErrorCode := 9;             // 非法状态兜底
    _eState := eFault;
END_CASE;

// ---- 完成标志统一出口映射 ----
xOpenDone := (_eState = eReady);
xCloseDone := (_eState = eDone);
eStateOut := _eState;
END_FUNCTION_BLOCK

(* ---- FB_DL_ServoDisableSafeSeq.st ---- *)
(* ===========================================================================
   组件名   : FB_DL_ServoDisableSafeSeq
   分类     : DL_Motion / 伺服安全下使能时序
   一句话   : 先减速到零速→撤使能→确认抱闸夹紧的安全下使能时序，任一步超时转故障态
   复杂度   : 1        版本 : v1.0.0        日期 : 2026-11-24
   开源溯源 : 无（clean-room 自研，未借鉴任何开源实现）
   输入契约 : xDisableReq 下使能请求；fVelAbs 速度绝对值 [rpm]；fZeroBand 零速带 [rpm]
              xEnableFbk 驱动器使能反馈；xBrakeClosedFbk 抱闸夹紧反馈
    工况边界  : 本件为「SS1 型受控停车序」（IEC 60204-1 停止类别 1 语义）：
                减速到零 -> 保持使能撤除 -> 抱闸闭合。适用于水平轴 / 无重力负载轴。
                **重力负载轴（垂直 Z 轴、举升轴）请改用 FB_DL_AxisBrakeSeq**：
                该件为抱闸优先序（先合抱闸建立力矩再撤使能），防自由滑落。
                二者顺序相反是工况差异所致，非缺陷；属主边界以本声明为准。
              t*Timeout 三步超时；xReset 复位上升沿
   输出契约 : xDecelCmd 减速指令；xEnableCmd 使能指令（撤使能后为 FALSE）
              xBrakeReleaseCmd 恒为 FALSE（失电夹紧为安全侧）
              xDone 时序完成；xError 故障锁存；iErrorCode 1=减速超时 2=撤使能超时
              3=抱闸超时 9=非法状态
   修改记录 : v1.0.0 2026-11-24 初版
   =========================================================================== *)

TYPE E_DL_DisableSeqState :
(
    eIdle := 0,          // 空闲 | idle
    eDecel := 1,         // 下发减速 | issue deceleration
    eWaitZero := 2,      // 等待零速 | wait zero speed
    eDisable := 3,       // 撤销使能 | drop enable
    eWaitDisable := 4,   // 等待使能撤销确认 | wait enable dropped
    eBrake := 5,         // 下发抱闸夹紧 | issue brake clamp
    eWaitBrake := 6,     // 等待抱闸确认 | wait brake confirm
    eDone := 7,          // 时序完成 | sequence done
    eFault := 8          // 故障锁存态 | latched fault
);
END_TYPE

FUNCTION_BLOCK FB_DL_ServoDisableSafeSeq
VAR_INPUT
    xDisableReq : BOOL;                     // 下使能请求 | disable request
    fVelAbs : REAL;                         // 速度绝对值 [rpm] | absolute speed [rpm]
    fZeroBand : REAL := 5.0;                // 零速判定带宽 [rpm] | zero speed band [rpm]
    xEnableFbk : BOOL;                      // 驱动器使能反馈 | drive enabled feedback
    xBrakeClosedFbk : BOOL;                 // 抱闸夹紧反馈 | brake clamped feedback
    tDecelTimeout : TIME := T#10S;          // 减速超时 | deceleration timeout
    tDisableTimeout : TIME := T#2S;         // 撤使能超时 | disable timeout
    tBrakeTimeout : TIME := T#2S;           // 抱闸夹紧超时 | brake timeout
    xReset : BOOL;                          // 故障复位上升沿 | fault reset rising edge
END_VAR
VAR_OUTPUT
    xDecelCmd : BOOL;                       // 减速指令 | deceleration command
    xEnableCmd : BOOL;                      // 使能指令 | enable command
    xBrakeReleaseCmd : BOOL;                // 抱闸释放指令（安全侧恒 FALSE） | brake release, always FALSE
    xDone : BOOL;                           // 时序完成 | sequence done
    xError : BOOL;                          // 故障锁存 | latched fault
    iErrorCode : INT;                       // 故障码 0=无故障 | error code
    eStateOut : E_DL_DisableSeqState;       // 当前状态观测 | current state observation
END_VAR
VAR
    _eState : E_DL_DisableSeqState := eIdle;  // 内部状态机状态 | internal state
    _xBadVel : BOOL;                      // 速度非有限或带宽非法 | velocity invalid
    _tonDecel : TON;                      // 减速等待定时器 | deceleration wait timer
    _tonDisable : TON;                    // 撤使能等待定时器 | disable wait timer
    _tonBrake : TON;                      // 抱闸等待定时器 | brake wait timer
    _rtReset : R_TRIG;                    // 复位上升沿 | reset rising edge
END_VAR

// ---- 速度合法性：非有限或带宽非正时视为未达零速 ----
_xBadVel := (fVelAbs <> fVelAbs) OR ((fVelAbs - fVelAbs) <> (fVelAbs - fVelAbs)) OR (fZeroBand <= 0.0);

// ---- 定时器与边沿：无条件每周期调用 ----
_tonDecel(IN := (_eState = eWaitZero), PT := tDecelTimeout);
_tonDisable(IN := (_eState = eWaitDisable), PT := tDisableTimeout);
_tonBrake(IN := (_eState = eWaitBrake), PT := tBrakeTimeout);
_rtReset(CLK := xReset);

// ---- 逐拍输出预置：非锁存量复位；抱闸释放恒 FALSE 为安全侧 ----
xDecelCmd := FALSE;
xEnableCmd := FALSE;
xBrakeReleaseCmd := FALSE;
xDone := FALSE;

CASE _eState OF
    eIdle:
        IF xDisableReq AND NOT xError THEN
            _eState := eDecel;
        END_IF

    eDecel:
        xDecelCmd := TRUE;
        xEnableCmd := TRUE;                      // 减速段必须保持使能，否则失控滑行
        _eState := eWaitZero;

    eWaitZero:
        xDecelCmd := TRUE;
        xEnableCmd := TRUE;
        IF (NOT _xBadVel) AND (ABS(fVelAbs) < fZeroBand) THEN
            _eState := eDisable;                 // 已到零速，可撤使能
        ELSIF _tonDecel.Q THEN
            xError := TRUE; iErrorCode := 1;     // 减速超时
            _eState := eFault;
        END_IF

    eDisable:
        _eState := eWaitDisable;                 // 本拍起使能指令保持 FALSE

    eWaitDisable:
        IF NOT xEnableFbk THEN
            _eState := eBrake;                   // 使能已撤销，再动抱闸
        ELSIF _tonDisable.Q THEN
            xError := TRUE; iErrorCode := 2;     // 撤使能超时
            _eState := eFault;
        END_IF

    eBrake:
        _eState := eWaitBrake;                   // 抱闸释放指令保持 FALSE，失电夹紧

    eWaitBrake:
        IF xBrakeClosedFbk THEN
            _eState := eDone;
        ELSIF _tonBrake.Q THEN
            xError := TRUE; iErrorCode := 3;     // 抱闸夹紧超时
            _eState := eFault;
        END_IF

    eDone:
        xDone := TRUE;
        IF NOT xDisableReq THEN
            _eState := eIdle;                    // 请求撤销后回空闲
        END_IF

    eFault:
        xError := TRUE;                          // 故障锁存保持，输出维持安全侧
        IF _rtReset.Q AND NOT xDisableReq THEN
            xError := FALSE;                     // 唯一解除路径：复位沿且无请求
            iErrorCode := 0;
            _eState := eIdle;
        END_IF

ELSE
    xError := TRUE; iErrorCode := 9;             // 非法状态兜底
    _eState := eFault;
END_CASE;

eStateOut := _eState;
END_FUNCTION_BLOCK

(* ---- FB_DL_ServoFollowErrMon.st ---- *)
(* ===========================================================================
   组件名   : FB_DL_ServoFollowErrMon
   分类     : DL_Motion / 伺服跟随误差监控
   一句话   : 位置指令与反馈之差经一阶低通后按预警/停机两级阈值分级报警，含非有限值拦截
   复杂度   : 2        版本 : v1.0.0        日期 : 2026-11-24
   开源溯源 : 无（clean-room 自研，未借鉴任何开源实现）
   输入契约 : xEnable 监控使能；lrPosCmd / lrPosFbk 位置指令与反馈 [mm]
              lrWarnLimit / lrStopLimit 两级阈值 [mm]；fLpfAlpha 低通系数 0..1
              tTripDelay 停机确认延时；xReset 复位上升沿
   输出契约 : lrFollowErr 滤波后跟随误差 [mm]；xWarn 预警（每拍重算，信息级）
              xStopTrip 停机锁存（唯一解除路径 = xReset 上升沿 AND 监控未使能）
              xValid 输入有效；iErrorCode 0=正常 1=输入非有限 2=阈值非法
   修改记录 : v1.0.0 2026-11-24 初版
   =========================================================================== *)

FUNCTION_BLOCK FB_DL_ServoFollowErrMon
VAR_INPUT
    xEnable : BOOL;                     // 监控使能 | monitoring enable
    lrPosCmd : LREAL;                   // 位置指令 [mm] | position command [mm]
    lrPosFbk : LREAL;                   // 位置反馈 [mm] | position feedback [mm]
    lrWarnLimit : LREAL := 5.0;         // 预警阈值 [mm] | warning limit [mm]
    lrStopLimit : LREAL := 10.0;        // 停机阈值 [mm] | stop limit [mm]
    fLpfAlpha : LREAL := 0.2;           // 一阶低通系数 0..1 | first order lpf alpha
    tTripDelay : TIME := T#50MS;        // 停机确认延时 | trip confirm delay
    xReset : BOOL;                      // 故障复位上升沿 | fault reset rising edge
END_VAR
VAR_OUTPUT
    lrFollowErr : LREAL;                // 滤波后跟随误差 [mm] | filtered following error [mm]
    xWarn : BOOL;                       // 预警输出（每拍重算） | warning output recomputed
    xStopTrip : BOOL;                   // 停机锁存输出 | latched stop trip
    xValid : BOOL;                      // 输入有效标志 | inputs valid flag
    iErrorCode : INT;                   // 故障码 0=无故障 | error code
END_VAR
VAR
    _lrErrMag : LREAL;                  // 误差绝对值 [mm] | absolute error [mm]
    _lrAlpha : LREAL;                   // 钳位后低通系数 | clamped lpf alpha
    _xBadCmd : BOOL;                    // 指令非有限 | command not finite
    _xBadFbk : BOOL;                    // 反馈非有限 | feedback not finite
    _xBadLim : BOOL;                    // 阈值非有限 | limits not finite
    _tonTrip : TON;                     // 停机确认定时器 | trip confirm timer
    _rtReset : R_TRIG;                  // 复位上升沿 | reset rising edge
END_VAR

// ---- 无条件每周期调用：复位沿检测 ----
_rtReset(CLK := xReset);

// ---- 非有限检测：NaN 用自反比较，Inf 用 (x-x)<>(x-x) ----
_xBadCmd := (lrPosCmd <> lrPosCmd) OR ((lrPosCmd - lrPosCmd) <> (lrPosCmd - lrPosCmd));
_xBadFbk := (lrPosFbk <> lrPosFbk) OR ((lrPosFbk - lrPosFbk) <> (lrPosFbk - lrPosFbk));
_xBadLim := (lrWarnLimit <> lrWarnLimit) OR ((lrWarnLimit - lrWarnLimit) <> (lrWarnLimit - lrWarnLimit))
         OR (lrStopLimit <> lrStopLimit) OR ((lrStopLimit - lrStopLimit) <> (lrStopLimit - lrStopLimit));

xValid := NOT (_xBadCmd OR _xBadFbk OR _xBadLim);
xWarn := FALSE;
iErrorCode := 0;
IF _xBadLim THEN
    iErrorCode := 2;                                  // 阈值非有限
ELSIF _xBadCmd OR _xBadFbk THEN
    iErrorCode := 1;                                  // 位置量非有限
END_IF
IF xValid AND ((lrWarnLimit <= 0.0) OR (lrStopLimit <= lrWarnLimit)) THEN
    xValid := FALSE;                                  // 阈值须为正值且停机阈值大于预警阈值
    iErrorCode := 2;
END_IF

// ---- 一阶低通：系数钳位到 0..1，避免发散 ----
_lrAlpha := fLpfAlpha;
IF _lrAlpha < 0.0 THEN
    _lrAlpha := 0.0;
ELSIF _lrAlpha > 1.0 THEN
    _lrAlpha := 1.0;
END_IF
IF xValid THEN
    _lrErrMag := ABS(lrPosCmd - lrPosFbk);
    lrFollowErr := lrFollowErr + _lrAlpha * (_lrErrMag - lrFollowErr);
ELSE
    lrFollowErr := 0.0;                               // 非法输入不污染滤波器状态
END_IF

// ---- 停机确认定时器：无条件每周期调用 ----
_tonTrip(IN := (lrFollowErr > lrStopLimit) AND xValid, PT := tTripDelay);

// ---- 两级分级判定 ----
xWarn := xValid AND (lrFollowErr > lrWarnLimit);
IF _tonTrip.Q THEN
    xStopTrip := TRUE;                                // 超阈值持续到延时后锁存
END_IF
IF _rtReset.Q AND NOT xEnable THEN
    xStopTrip := FALSE;                               // 唯一解除路径：复位沿且监控未使能
END_IF
IF NOT xEnable THEN
    xWarn := FALSE;                                   // 未使能时预警不对外输出
END_IF
END_FUNCTION_BLOCK

(* ---- FB_DL_ServoOverloadDerate.st ---- *)
(* ===========================================================================
   组件名   : FB_DL_ServoOverloadDerate
   分类     : DL_Motion / 伺服过载降额
   一句话   : 按连续负载率与 I2t 累积量计算转矩降额系数，恢复时带滞回并锁存过载报警
   复杂度   : 2        版本 : v1.0.0        日期 : 2026-11-24
   开源溯源 : 无（clean-room 自研，未借鉴任何开源实现）
   输入契约 : xEnable 功能使能；fLoadRatio 连续负载率 1.0=额定；fDtSec 采样周期 [s]
              fI2tLimit 累积限值 [%·s]；fCoolGain 冷却泄放增益 [1/s]
              fDerateStart 降额起始负载率；fDerateMin 最小降额系数；fHyst 恢复滞回带
              xReset 过载锁存复位沿
   输出契约 : fDerateFactor 降额系数 0..1；fI2tAccum 累积量 [%·s]
              xDerated 降额生效（滞回保持）；xOverload 过载锁存
              xValid 输入有效；iErrorCode 0=正常 1=非有限 2=参数非法 3=过载
   修改记录 : v1.0.0 2026-11-24 初版
   =========================================================================== *)

FUNCTION_BLOCK FB_DL_ServoOverloadDerate
VAR_INPUT
    xEnable : BOOL;                     // 降额功能使能 | derating enable
    fLoadRatio : REAL;                  // 连续负载率 1.0=额定 | continuous load ratio
    fDtSec : REAL := 0.004;             // 采样周期 [s] | sample period [s]
    fI2tLimit : REAL := 100.0;          // I2t 累积限值 [%·s] | i2t limit [%·s]
    fCoolGain : REAL := 1.0;            // 冷却泄放增益 [1/s] | cooling decay gain [1/s]
    fDerateStart : REAL := 0.8;         // 降额起始负载率 | derate start ratio
    fDerateMin : REAL := 0.3;           // 最小降额系数 | minimum derate factor
    fHyst : REAL := 0.05;               // 恢复滞回带宽 | recovery hysteresis band
    xReset : BOOL;                      // 过载锁存复位沿 | overload reset edge
END_VAR
VAR_OUTPUT
    fDerateFactor : REAL;               // 转矩降额系数 0..1 | torque derate factor
    fI2tAccum : REAL;                   // I2t 累积量 [%·s] | i2t accumulator [%·s]
    xDerated : BOOL;                    // 降额生效标志（滞回） | derating active with hysteresis
    xOverload : BOOL;                   // 过载锁存报警 | latched overload alarm
    xValid : BOOL;                      // 输入有效标志 | inputs valid flag
    iErrorCode : INT;                   // 故障码 0=无故障 | error code
END_VAR
VAR
    _fDt : REAL;                        // 钳位后采样周期 [s] | clamped dt [s]
    _fR : REAL;                         // 钳位后负载率 | clamped load ratio
    _fI2t : REAL;                       // 内部 I2t 累积量 [%·s] | internal i2t accumulator
    _fDen : REAL;                       // 降额计算分母 | derate denominator
    _xBad : BOOL;                       // 输入非有限标志 | not-finite flag
    _xBadPar : BOOL;                    // 参数非法标志 | invalid parameter flag
    _rtReset : R_TRIG;                  // 复位上升沿 | reset rising edge
END_VAR

// ---- 无条件每周期调用：复位沿检测 ----
_rtReset(CLK := xReset);

// ---- 非有限值检测 ----
_xBad := (fLoadRatio <> fLoadRatio) OR ((fLoadRatio - fLoadRatio) <> (fLoadRatio - fLoadRatio))
      OR (fDtSec <> fDtSec) OR ((fDtSec - fDtSec) <> (fDtSec - fDtSec))
      OR (fI2tLimit <> fI2tLimit) OR ((fI2tLimit - fI2tLimit) <> (fI2tLimit - fI2tLimit))
      OR (fCoolGain <> fCoolGain) OR ((fCoolGain - fCoolGain) <> (fCoolGain - fCoolGain));

// ---- 参数合法性：所有分母与滞回带必须为正 ----
_xBadPar := (fI2tLimit <= 0.0) OR (fCoolGain <= 0.0) OR (fHyst < 0.0)
         OR (fDerateStart <= 0.0) OR (fDerateStart >= 1.0)
         OR (fDerateMin <= 0.0) OR (fDerateMin >= 1.0);

// ---- 输出预置：xDerated / xOverload 为保持量，不在本处清零 ----
fDerateFactor := 1.0;
xValid := FALSE;
iErrorCode := 0;
IF _xBad THEN
    iErrorCode := 1;                                  // 输入非有限
ELSIF _xBadPar THEN
    iErrorCode := 2;                                  // 参数非法
END_IF

IF _xBad OR _xBadPar THEN
    fDerateFactor := 1.0;                             // 参数不可信时保守输出满转矩
    fI2tAccum := _fI2t;
ELSE
    xValid := TRUE;

    // 周期钳位：防止零除与超大积分步长
    _fDt := fDtSec;
    IF _fDt < 0.000001 THEN
        _fDt := 0.000001;
    ELSIF _fDt > 0.2 THEN
        _fDt := 0.2;
    END_IF
    _fR := fLoadRatio;
    IF _fR < 0.0 THEN
        _fR := 0.0;
    ELSIF _fR > 10.0 THEN
        _fR := 10.0;
    END_IF

    // ---- I2t 累积与冷却泄放 ----
    IF _fR > 1.0 THEN
        _fI2t := _fI2t + (_fR * _fR - 1.0) * _fDt;    // 过载段净累积
    ELSE
        _fI2t := _fI2t - fCoolGain * (1.0 - _fR) * _fDt;  // 轻载段泄放
    END_IF
    IF _fI2t < 0.0 THEN
        _fI2t := 0.0;                                 // 累积量不取负值
    END_IF

    // ---- 滞回判定降额生效：进入无滞回，退出需低于起始值且累积已泄完 ----
    IF _fR >= fDerateStart THEN
        xDerated := TRUE;
    ELSIF (_fR < (fDerateStart - fHyst)) AND (_fI2t <= 0.0) THEN
        xDerated := FALSE;
    END_IF

    // ---- 降额系数：起始负载率到额定线性过渡 ----
    IF xDerated THEN
        _fDen := 1.0 - fDerateStart;
        IF _fDen > 0.000000001 THEN
            fDerateFactor := 1.0 - (1.0 - fDerateMin) * (_fR - fDerateStart) / _fDen;
        END_IF
        IF fDerateFactor < fDerateMin THEN
            fDerateFactor := fDerateMin;
        ELSIF fDerateFactor > 1.0 THEN
            fDerateFactor := 1.0;
        END_IF
    END_IF

    // ---- 过载锁存与唯一解除路径 ----
    IF _fI2t >= fI2tLimit THEN
        xOverload := TRUE;
    END_IF
    IF _rtReset.Q AND NOT xEnable THEN
        xOverload := FALSE;                           // 解除路径：复位沿且功能未使能
        _fI2t := 0.0;
    END_IF
    IF xOverload THEN
        iErrorCode := 3;                              // 过载锁存状态优先
    END_IF
    fI2tAccum := _fI2t;
END_IF
END_FUNCTION_BLOCK

(* ---- FB_DL_ServoRegenEnergyCalc.st ---- *)
(* ===========================================================================
   组件名   : FB_DL_ServoRegenEnergyCalc
   分类     : DL_Motion / 伺服再生能耗估算
   一句话   : 由减速段动能差与回馈效率估算再生功率与累积能量，超限锁存报警
   复杂度   : 2        版本 : v1.0.0        日期 : 2026-11-24
   开源溯源 : 无（clean-room 自研，未借鉴任何开源实现）
   输入契约 : xEnable 功能使能；fInertia 折算惯量 [kg·m²]；fVelNowRad 当前角速度 [rad/s]
              fDtSec 采样周期 [s]；fEfficiency 回馈效率 0..1；fEnergyLimitWh 累积限值 [Wh]
              xReset 超限锁存复位沿
   输出契约 : fRegenPowerW 本拍再生功率 [W]；fEnergyAccumWh 累积再生能量 [Wh]
              fKineticJ 本拍动能 [J]；xRegenActive 处于再生（减速）段
              xOverLimit 累积超限锁存；xValid 输入有效
              iErrorCode 0=正常 1=非有限 2=参数非法 3=累积超限
   修改记录 : v1.0.0 2026-11-24 初版
   =========================================================================== *)

FUNCTION_BLOCK FB_DL_ServoRegenEnergyCalc
VAR_INPUT
    xEnable : BOOL;                     // 功能使能 | function enable
    fInertia : REAL := 0.001;           // 折算惯量 [kg·m²] | reflected inertia [kg·m²]
    fVelNowRad : REAL;                  // 当前角速度 [rad/s] | current angular velocity [rad/s]
    fDtSec : REAL := 0.004;             // 采样周期 [s] | sample period [s]
    fEfficiency : REAL := 0.85;         // 回馈效率 0..1 | regen efficiency 0..1
    fEnergyLimitWh : REAL := 50.0;      // 累积能量限值 [Wh] | energy limit [Wh]
    xReset : BOOL;                      // 超限锁存复位沿 | over-limit reset edge
END_VAR
VAR_OUTPUT
    fRegenPowerW : REAL;                // 本拍再生功率 [W] | regen power this cycle [W]
    fEnergyAccumWh : REAL;              // 累积再生能量 [Wh] | accumulated regen energy [Wh]
    fKineticJ : REAL;                   // 本拍旋转动能 [J] | kinetic energy [J]
    xRegenActive : BOOL;                // 处于再生段 | regeneration active
    xOverLimit : BOOL;                  // 累积超限锁存 | latched over-limit
    xValid : BOOL;                      // 输入有效标志 | inputs valid flag
    iErrorCode : INT;                   // 故障码 0=无故障 | error code
END_VAR
VAR
    _fKePrev : REAL;                    // 上一拍动能 [J] | previous kinetic energy [J]
    _fKeNow : REAL;                     // 本拍动能 [J] | current kinetic energy [J]
    _fDeltaJ : REAL;                    // 动能差 [J] | kinetic energy difference [J]
    _fDt : REAL;                        // 钳位后采样周期 [s] | clamped dt [s]
    _fAccum : REAL;                     // 内部累积能量 [Wh] | internal accumulator [Wh]
    _xBad : BOOL;                       // 输入非有限标志 | not-finite flag
    _xBadPar : BOOL;                    // 参数非法标志 | invalid parameter flag
    _rtReset : R_TRIG;                  // 复位上升沿 | reset rising edge
END_VAR

// ---- 无条件每周期调用：复位沿检测 ----
_rtReset(CLK := xReset);

// ---- 非有限检测 ----
_xBad := (fInertia <> fInertia) OR ((fInertia - fInertia) <> (fInertia - fInertia))
      OR (fVelNowRad <> fVelNowRad) OR ((fVelNowRad - fVelNowRad) <> (fVelNowRad - fVelNowRad))
      OR (fDtSec <> fDtSec) OR ((fDtSec - fDtSec) <> (fDtSec - fDtSec))
      OR (fEfficiency <> fEfficiency) OR ((fEfficiency - fEfficiency) <> (fEfficiency - fEfficiency));

// ---- 参数合法性：惯量非负、效率落在 (0,1]、限值为正 ----
_xBadPar := (fInertia < 0.0) OR (fEfficiency <= 0.0) OR (fEfficiency > 1.0)
         OR (fEnergyLimitWh <= 0.0) OR (fDtSec <= 0.0);

// ---- 输出预置 ----
fRegenPowerW := 0.0;
fKineticJ := 0.0;
xRegenActive := FALSE;
xValid := NOT (_xBad OR _xBadPar);
iErrorCode := 0;
IF _xBad THEN
    iErrorCode := 1;
ELSIF _xBadPar THEN
    iErrorCode := 2;
END_IF

// ---- 周期钳位：防零除与超大积分步长 ----
_fDt := fDtSec;
IF _fDt < 0.000001 THEN
    _fDt := 0.000001;
ELSIF _fDt > 0.2 THEN
    _fDt := 0.2;
END_IF

IF xValid AND xEnable THEN
    // ---- 动能计算：Ek = 0.5 * J * w^2 ----
    _fKeNow := 0.5 * fInertia * fVelNowRad * fVelNowRad;
    fKineticJ := _fKeNow;

    // ---- 再生判定：仅当本拍动能低于上拍（减速）才有能量回馈 ----
    _fDeltaJ := _fKePrev - _fKeNow;
    IF _fDeltaJ > 0.0 THEN
        xRegenActive := TRUE;
        fRegenPowerW := _fDeltaJ / _fDt * fEfficiency;        // 分母已守卫
        _fAccum := _fAccum + _fDeltaJ * fEfficiency / 3600.0;  // J -> Wh
    END_IF

    // ---- 超限置位 ----
    IF _fAccum >= fEnergyLimitWh THEN
        xOverLimit := TRUE;
    END_IF

    // ---- 状态推进：动能快照留到拍末生效 ----
    _fKePrev := _fKeNow;
END_IF

// ---- 超限锁存与唯一解除路径 ----
// 解除门要求 NOT xEnable，必须放在使能门控块之外评估，否则该路径永不可达
IF _rtReset.Q AND NOT xEnable THEN
    xOverLimit := FALSE;
    _fAccum := 0.0;
END_IF
IF xOverLimit THEN
    iErrorCode := 3;                                      // 超限锁存状态优先
END_IF

fEnergyAccumWh := _fAccum;
END_FUNCTION_BLOCK

(* ---- FB_DL_ServoStiffnessSwitch.st ---- *)
(* ===========================================================================
   组件名   : FB_DL_ServoStiffnessSwitch
   分类     : DL_Motion / 伺服刚性档位
   一句话   : 静止/低速/高速三档增益组切换，切换须零速且增益按斜坡过渡，禁止带速硬切
   复杂度   : 2        版本 : v1.0.0        日期 : 2026-11-24
   开源溯源 : 无（clean-room 自研，未借鉴任何开源实现）
   输入契约 : xEnable 功能使能；eGearReq 目标档位请求；fVelAbs 当前速度绝对值 [rpm]
              fZeroSpeedBand 零速判定带宽 [rpm]；afKp/afKi/afKd 三档增益表 [1..3]
              fRampRate 增益过渡速率 [1/s]；fDtSec 采样周期 [s]
   输出契约 : fKpAct/fKiAct/fKdAct 生效增益；eGearAct 生效档位；xSwitchBusy 过渡中
              xSwitchBlocked 因速度过高被拒切换；xValid 输入有效
              iErrorCode 0=正常 1=非有限 2=参数非法 9=非法档位
   修改记录 : v1.0.0 2026-11-24 初版
   =========================================================================== *)

TYPE E_DL_StiffGear :
(
    eStaticGain := 0,    // 静止高刚性档 | standstill high stiffness
    eLowSpeedGain := 1,  // 低速中刚性档 | low speed medium stiffness
    eHighSpeedGain := 2  // 高速低刚性档 | high speed low stiffness
);
END_TYPE

FUNCTION_BLOCK FB_DL_ServoStiffnessSwitch
VAR_INPUT
    xEnable : BOOL;                             // 功能使能 | function enable
    eGearReq : E_DL_StiffGear := eStaticGain;   // 目标档位请求 | requested gear
    fVelAbs : REAL;                             // 速度绝对值 [rpm] | absolute speed [rpm]
    fZeroSpeedBand : REAL := 5.0;               // 零速判定带宽 [rpm] | zero speed band [rpm]
    afKp : ARRAY[1..3] OF REAL;                 // 三档比例增益表 | three gear kp table
    afKi : ARRAY[1..3] OF REAL;                 // 三档积分增益表 | three gear ki table
    afKd : ARRAY[1..3] OF REAL;                 // 三档微分增益表 | three gear kd table
    fRampRate : REAL := 20.0;                   // 增益过渡速率 [1/s] | gain ramp rate [1/s]
    fDtSec : REAL := 0.004;                     // 采样周期 [s] | sample period [s]
END_VAR
VAR_OUTPUT
    fKpAct : REAL;                              // 生效比例增益 | active kp
    fKiAct : REAL;                              // 生效积分增益 | active ki
    fKdAct : REAL;                              // 生效微分增益 | active kd
    eGearAct : E_DL_StiffGear;                  // 生效档位（默认首项=静止档） | active gear
    xSwitchBusy : BOOL;                         // 增益过渡进行中 | gain ramp in progress
    xSwitchBlocked : BOOL;                      // 带速切换被拒 | switch rejected at speed
    xValid : BOOL;                              // 输入有效标志 | inputs valid flag
    iErrorCode : INT;                           // 故障码 0=无故障 | error code
END_VAR
VAR
    _iIdxAct : INT := 1;                        // 生效档位数组下标 1..3 | active index
    _iIdxReq : INT := 1;                        // 请求档位数组下标 1..3 | requested index
    _i : INT := 1;                              // 循环下标 | loop index
    _fDt : REAL;                                // 钳位后采样周期 [s] | clamped dt [s]
    _fStep : REAL;                              // 单拍增益步长 | gain step per cycle
    _afAct : ARRAY[1..3] OF REAL;               // 当前生效增益缓存 | active gain buffer
    _afTgt : ARRAY[1..3] OF REAL;               // 目标增益缓存 | target gain buffer
    _xBad : BOOL;                               // 输入非有限标志 | not-finite flag
    _xBadPar : BOOL;                            // 参数非法标志 | invalid parameter flag
END_VAR

// ---- 非有限检测 ----
_xBad := (fVelAbs <> fVelAbs) OR ((fVelAbs - fVelAbs) <> (fVelAbs - fVelAbs))
      OR (fRampRate <> fRampRate) OR ((fRampRate - fRampRate) <> (fRampRate - fRampRate))
      OR (fDtSec <> fDtSec) OR ((fDtSec - fDtSec) <> (fDtSec - fDtSec));
_i := 1;
WHILE _i <= 3 DO
    IF ((afKp[_i] <> afKp[_i]) OR (afKi[_i] <> afKi[_i]) OR (afKd[_i] <> afKd[_i])) THEN
        _xBad := TRUE;                          // 任一档增益非有限即判无效
    END_IF
    _i := _i + 1;
END_WHILE

// ---- 参数合法性 ----
_xBadPar := (fZeroSpeedBand <= 0.0) OR (fRampRate <= 0.0) OR (fDtSec <= 0.0);

// ---- 输出预置：非锁存量复位 ----
xSwitchBusy := FALSE;
xSwitchBlocked := FALSE;
xValid := NOT (_xBad OR _xBadPar);
iErrorCode := 0;
IF _xBad THEN
    iErrorCode := 1;
ELSIF _xBadPar THEN
    iErrorCode := 2;
END_IF

// ---- 档位到数组下标映射：禁止枚举直接转型，用 CASE 显式映射 ----
CASE eGearAct OF
    eStaticGain: _iIdxAct := 1;
    eLowSpeedGain: _iIdxAct := 2;
    eHighSpeedGain: _iIdxAct := 3;
ELSE
    _iIdxAct := 1;                              // 非法生效档位兜底回静止档
    iErrorCode := 9;
END_CASE
CASE eGearReq OF
    eStaticGain: _iIdxReq := 1;
    eLowSpeedGain: _iIdxReq := 2;
    eHighSpeedGain: _iIdxReq := 3;
ELSE
    _iIdxReq := 1;                              // 非法请求档位兜底回静止档
    iErrorCode := 9;
END_CASE
IF _iIdxAct < 1 THEN
    _iIdxAct := 1;
ELSIF _iIdxAct > 3 THEN
    _iIdxAct := 3;
END_IF
IF _iIdxReq < 1 THEN
    _iIdxReq := 1;
ELSIF _iIdxReq > 3 THEN
    _iIdxReq := 3;
END_IF

// ---- 切换许可：须功能使能且零速，否则拒绝并置阻塞标志 ----
IF (_iIdxReq <> _iIdxAct) AND xValid AND xEnable THEN
    IF ABS(fVelAbs) < fZeroSpeedBand THEN
        eGearAct := eGearReq;                   // 零速许可切换
        _iIdxAct := _iIdxReq;
    ELSE
        xSwitchBlocked := TRUE;                 // 带速切换被拒，保持原档
    END_IF
END_IF

// ---- 增益斜坡过渡（受使能与合法性门控） ----
_fDt := fDtSec;
IF _fDt > 0.2 THEN
    _fDt := 0.2;                                // 周期上限，防大步长跳变
END_IF
_fStep := fRampRate * _fDt;
IF NOT xValid THEN
    _fStep := 0.0;                              // 非法输入时冻结过渡
END_IF

_afAct[1] := fKpAct;
_afAct[2] := fKiAct;
_afAct[3] := fKdAct;
_afTgt[1] := afKp[_iIdxAct];
_afTgt[2] := afKi[_iIdxAct];
_afTgt[3] := afKd[_iIdxAct];

FOR _i := 1 TO 3 DO
    IF _afAct[_i] < _afTgt[_i] THEN
        _afAct[_i] := _afAct[_i] + _fStep;
        IF _afAct[_i] > _afTgt[_i] THEN
            _afAct[_i] := _afTgt[_i];
        END_IF
    ELSIF _afAct[_i] > _afTgt[_i] THEN
        _afAct[_i] := _afAct[_i] - _fStep;
        IF _afAct[_i] < _afTgt[_i] THEN
            _afAct[_i] := _afTgt[_i];
        END_IF
    END_IF
END_FOR

// ---- 过渡完成判定：三路增益均已收敛（用容差比较，禁止浮点等值） ----
xSwitchBusy := (ABS(_afAct[1] - _afTgt[1]) > 0.000000001)
            OR (ABS(_afAct[2] - _afTgt[2]) > 0.000000001)
            OR (ABS(_afAct[3] - _afTgt[3]) > 0.000000001);

fKpAct := _afAct[1];
fKiAct := _afAct[2];
fKdAct := _afAct[3];
IF NOT xEnable THEN
    xSwitchBlocked := FALSE;                    // 未使能时不上报阻塞
END_IF
END_FUNCTION_BLOCK

(* ---- FB_DL_ServoTorqueClamp.st ---- *)
(* ===========================================================================
   组件名   : FB_DL_ServoTorqueClamp
   分类     : DL_Motion / 伺服转矩限幅
   一句话   : 按工艺段查表得正负转矩上限，再按电机温度线性降额，输出限幅生效标志
   复杂度   : 2        版本 : v1.0.0        日期 : 2026-11-24
   开源溯源 : 无（clean-room 自研，未借鉴任何开源实现）
   输入契约 : eSeg 工艺段；afPosLim/afNegLim 五段正负转矩上限表 [%]（按段号 1..5）
              fTempMotor 电机温度 [°C]；fTempDerateStart 降额起始温度 [°C]
              fTempDerateEnd 降额终止温度 [°C]；fDerateFloor 最低降额系数
   输出契约 : fTorqueLimPos 正向转矩上限 [%]；fTorqueLimNeg 反向转矩上限（负值）[%]
              fDerateFactor 温度降额系数 0..1；xClampActive 限幅生效（降额<1）
              xValid 输入有效；iErrorCode 0=正常 1=非有限 2=参数非法 9=非法段号
   修改记录 : v1.0.0 2026-11-24 初版
   =========================================================================== *)

TYPE E_DL_TorqueSeg :
(
    eSegIdle := 0,   // 空闲段 | idle segment
    eSegAccel := 1,  // 加速段 | acceleration segment
    eSegRun := 2,    // 匀速段 | constant speed segment
    eSegDecel := 3,  // 减速段 | deceleration segment
    eSegHold := 4    // 保持段 | holding segment
);
END_TYPE

FUNCTION_BLOCK FB_DL_ServoTorqueClamp
VAR_INPUT
    eSeg : E_DL_TorqueSeg := eSegIdle;      // 当前工艺段 | current process segment
    afPosLim : ARRAY[1..5] OF REAL;         // 五段正向转矩上限 [%] | positive limits [%]
    afNegLim : ARRAY[1..5] OF REAL;         // 五段反向转矩上限 [%] | negative limits [%]
    fTempMotor : REAL := 25.0;              // 电机温度 [°C] | motor temperature [°C]
    fTempDerateStart : REAL := 60.0;        // 降额起始温度 [°C] | derate start temp [°C]
    fTempDerateEnd : REAL := 90.0;          // 降额终止温度 [°C] | derate end temp [°C]
    fDerateFloor : REAL := 0.2;             // 最低降额系数 | minimum derate factor
END_VAR
VAR_OUTPUT
    fTorqueLimPos : REAL;                   // 正向转矩上限 [%] | positive torque limit [%]
    fTorqueLimNeg : REAL;                   // 反向转矩上限（负值）[%] | negative torque limit [%]
    fDerateFactor : REAL;                   // 温度降额系数 0..1 | temperature derate factor
    xClampActive : BOOL;                    // 限幅生效标志 | clamp active flag
    xValid : BOOL;                          // 输入有效标志 | inputs valid flag
    iErrorCode : INT;                       // 故障码 0=无故障 | error code
END_VAR
VAR
    _iSeg : INT := 1;                       // 段号数组下标 1..5 | segment index 1..5
    _i : INT := 1;                          // 循环下标 | loop index
    _fPosBase : REAL;                       // 表内正向基值 [%] | table positive base [%]
    _fNegBase : REAL;                       // 表内反向基值 [%] | table negative base [%]
    _fSpan : REAL;                          // 温度降额区间宽度 [°C] | derate span [°C]
    _xBad : BOOL;                           // 输入非有限标志 | not-finite flag
    _xBadPar : BOOL;                        // 参数非法标志 | invalid parameter flag
END_VAR

// ---- 非有限检测 ----
_xBad := (fTempMotor <> fTempMotor) OR ((fTempMotor - fTempMotor) <> (fTempMotor - fTempMotor))
      OR (fTempDerateStart <> fTempDerateStart) OR ((fTempDerateStart - fTempDerateStart) <> (fTempDerateStart - fTempDerateStart))
      OR (fTempDerateEnd <> fTempDerateEnd) OR ((fTempDerateEnd - fTempDerateEnd) <> (fTempDerateEnd - fTempDerateEnd));
_i := 1;
WHILE _i <= 5 DO
    IF (afPosLim[_i] <> afPosLim[_i]) OR (afNegLim[_i] <> afNegLim[_i]) THEN
        _xBad := TRUE;                      // 表内任一项非有限即判无效
    END_IF
    _i := _i + 1;
END_WHILE

// ---- 参数合法性：降额区间必须正向有序，系数落在 0..1 ----
_fSpan := fTempDerateEnd - fTempDerateStart;
_xBadPar := (_fSpan <= 0.000000001) OR (fDerateFloor <= 0.0) OR (fDerateFloor > 1.0);

// ---- 输出预置 ----
fTorqueLimPos := 0.0;
fTorqueLimNeg := 0.0;
fDerateFactor := 1.0;
xClampActive := FALSE;
xValid := NOT (_xBad OR _xBadPar);
iErrorCode := 0;
IF _xBad THEN
    iErrorCode := 1;
ELSIF _xBadPar THEN
    iErrorCode := 2;
END_IF

// ---- 段号到数组下标映射：用 CASE 显式映射，禁止枚举直接转型 ----
CASE eSeg OF
    eSegIdle: _iSeg := 1;
    eSegAccel: _iSeg := 2;
    eSegRun: _iSeg := 3;
    eSegDecel: _iSeg := 4;
    eSegHold: _iSeg := 5;
ELSE
    _iSeg := 1;                             // 非法段号兜底回空闲段
    iErrorCode := 9;
END_CASE
IF _iSeg < 1 THEN
    _iSeg := 1;                             // 下标钳位，防越界
ELSIF _iSeg > 5 THEN
    _iSeg := 5;
END_IF

IF xValid THEN
    // ---- 温度降额：起始温度以下不降，终止温度以上压到地板值 ----
    IF fTempMotor <= fTempDerateStart THEN
        fDerateFactor := 1.0;
    ELSIF fTempMotor >= fTempDerateEnd THEN
        fDerateFactor := fDerateFloor;
    ELSE
        fDerateFactor := 1.0 - (1.0 - fDerateFloor) * (fTempMotor - fTempDerateStart) / _fSpan;
        IF fDerateFactor < fDerateFloor THEN
            fDerateFactor := fDerateFloor;
        ELSIF fDerateFactor > 1.0 THEN
            fDerateFactor := 1.0;
        END_IF
    END_IF

    // ---- 表值取绝对值作为幅值，正负号由输出方向分别表达 ----
    _fPosBase := ABS(afPosLim[_iSeg]);
    _fNegBase := ABS(afNegLim[_iSeg]);
    fTorqueLimPos := _fPosBase * fDerateFactor;
    fTorqueLimNeg := -_fNegBase * fDerateFactor;    // 反向限幅输出负值

    // ---- 限幅生效：降额系数明显小于 1 即为生效 ----
    xClampActive := (fDerateFactor < 0.999999999);
END_IF
// 非法输入分支不覆盖上限：预置的 0 转矩上限即为安全侧输出（禁止自赋值死语句）
END_FUNCTION_BLOCK
